(* IEC 61131-3 sources: daoli-st-library/DL_Base, 243 files *)

(* ---- E_DL_ControlModeSel.st ---- *)
// E_DL_ControlModeSel v1.0.0
// 开源溯源：AixOCAT / URL https://github.com/AixOCAT / 许可证 MIT / 借鉴 CONTROL_MODE 枚举语义（手/自动/停止三态），clean-room 重写
(*
  道莅工业代码库 | DL_Base | E_DL_ControlModeSel
  版本: 1.0.0 | 日期: 2026-11-23 | 轮次: R75
  功能: 手动/自动/停止三态控制模式枚举（strict 口径，配 MANUAL 覆写件族）
  邻件关系: 与 E_SMStatus 语义相邻（状态机状态 vs 操作模式选择），本件为
            模式选择属主；引用方（覆写/手自动切换族）只引用不重声明（R12）
  使用约定: 全库唯一属主，其他件引用时由 L2 闸按类型名自动回溯本文件；
            成员值固定步进 10，禁止中途插值改序（防历史引用漂移）
*)
TYPE E_DL_ControlModeSel :
(
    eManual := 0,    // 手动模式（操作员直控，联锁保留）/ Manual mode, operator direct with interlocks
    eAuto   := 10,   // 自动模式（程序/上位调度）/ Auto mode, program or supervisory driven
    eStop   := 20    // 停止模式（受控停机，输出回安全位）/ Stop mode, controlled stop to safe outputs
);
END_TYPE

(* ---- FB_DL_EStopMonitor.st ---- *)
(*==============================================================================
 * 组件名称 (Component)  : FB_DL_EStopMonitor
 * 所属子库 (Sublibrary) : DL_Base
 * 当前版本 (Version)    : 1.0.0
 * 兼容性   (Platform)   : CODESYS 3.5+ / TwinCAT 3 / 汇川 InoProShop / 施耐德 Machine Expert
 *                         仅依赖 Standard.library（TON / R_TRIG / F_TRIG / ABS），
 *                         零厂商私有库
 * 功能描述 (Function)   : 急停双通道监视：通道语义 TRUE=回路闭合（健康）。
 *                         任一通道断开 → bSafe 立即 FALSE（安全侧一级拦截，
 *                         不等确认窗）；两通道电平不一致（bCh1 <> bCh2）持续
 *                         tMismatchWin → bMismatch 锁存 + 首出通道号 eFirstOut
 *                         锁存（先断开的通道，F_TRIG 双实例竞争记录）；复位须
 *                         双通道恢复一致（bCh1 ∧ bCh2）且 bReset 上升沿才清
 *                         bMismatch/首出（规格指定）。
 * 接口     (Interface)  : 输入 bCh1 通道 1（TRUE=闭合健康）、bCh2 通道 2、
 *                         tMismatchWin 失配确认窗（域 > T#0S）、bReset 复位；
 *                         输出 bSafe 可运行判据（双通道健康 ∧ 无失配锁存）、
 *                         bMismatch 失配锁存、eFirstOut 首出通道号（锁存）、
 *                         eErrCode 错误码、bError 故障标志。
 * 边界     (Boundary)   : ① **属主边界（写死）：本件只做双通道监视判据，不切断
 *                         执行器、不做安全认证**（安全切断由安全继电器/IO 映射层
 *                         双保险执行，本件为诊断与允许运行判据源）。
 *                         ② 首出归因：双 F_TRIG 竞争窗口内先到沿者赢（同拍
 *                         双断时按 bCh1 优先判定，头注释声明：同拍双断无法区分
 *                         物理先后，eFirstOut 取 eCh1，规格允许的确定性归因）。
 *                         ③ 双通道同拍齐断（一致断开）不判失配：bSafe=FALSE
 *                         照常拦截，eFirstOut 保持 eNone（一致事件无失配语义）。
 *                         ④ 失配确认 TON 的 IN 派生式（bCh1 <> bCh2）∧ 通道
 *                         未齐断，段 0 无条件调用；出窗自复位（不一致消失即
 *                         复位，无外部沿清零依赖）。
 *                         ⑤ 锁存解除路径：bMismatch/eFirstOut 解除边 = 双通道
 *                         健康 ∧ bReset 上升沿（可达，头注释声明，R188/R152）。
 *                         ⑥ 零全局耦合（无 GVL / VAR_EXTERNAL / 物理地址）。
 * 分工声明 (Scope)      : 与 `FB_DL_RedundantSwitch` 分工：通道二选一归那件、
 *                         急停一致性监视归本件；与 `FB_DL_EdgeOrderCheck` 分工：
 *                         通用顺序校验归那件，本件首出归因为急停专用语义。
 * 来源标签 (Source Tag) : IEC 61131-3 标准语义的道莅防御性实现（双通道一致性
 *                         监视为标准安全监视语义）
 * 码表     (Codes)      : 本件不占用任何全局数字码位。出口为 BOOL 组 +
 *                         ENUM 通道号/错误码；数字码位待主控收口阶段统一派号。
 * 红线自检 (Redline)    : R1 ✓ 零 GVL/VAR_EXTERNAL ｜ R2 ✓ 零 %I/%Q/%M ｜ R3 ✓ 纯 IEC 61131-3
 *                         R4 ✓ 一级拦截不等窗 + 锁存解除可达 + 归因唯一 ｜ R5 ✓ 声明逐行同行双语注释
 *                         R6 ✓ ENUM 状态机不用（首出枚举 + 锁存态） ｜ R7 ✓ 一 TON 两 F_TRIG 一 R_TRIG 段 0 无条件刷新
 * 修订历史 (Revision)   : 2026-11-20  v1.0.0  R50 首版（批次 2 · 序号 10）
 * 验收向量 (Acceptance) : ① 双通道 TRUE，bCh1 在 t0 断开且 tMismatchWin 内未
 *                         恢复 → bMismatch=TRUE、eFirstOut=eCh1、bSafe=FALSE；
 *                         ② bCh1 断开 20ms 内恢复（tMismatchWin=100MS）→
 *                         tonMis 未到，bMismatch 保持 FALSE；③ 失配锁存后
 *                         bCh1/bCh2 均 TRUE + bReset 上升沿 → bMismatch=
 *                         FALSE、eFirstOut=eNone、bSafe=TRUE；④ 双通道同拍
 *                         齐断 → bSafe=FALSE，bMismatch=FALSE，eFirstOut=eNone。
 *==============================================================================*)

(*-----------------------------------------------------------------------------
 * 枚举: E_DL_EstChannel（首出通道号，锁存回放）
 *----------------------------------------------------------------------------*)
TYPE E_DL_EstChannel :
(
    eNone := 0,   // 无首出（未发生失配或同拍齐断） / No first-out
    eCh1  := 1,   // 首出通道 1 / First-out channel 1
    eCh2  := 2    // 首出通道 2 / First-out channel 2
);
END_TYPE

(*-----------------------------------------------------------------------------
 * 枚举: E_DL_EstErr（错误码；信息级不置 bError，故障级恒伴 bError=TRUE）
 *----------------------------------------------------------------------------*)
TYPE E_DL_EstErr :
(
    eOk      := 0,   // 正常 / Normal
    eCfgBad  := 1,   // 故障级：确认窗组态非法（<= T#0S） / Fault: window config illegal
    eMisLock := 2    // 故障级：失配锁存回放（归因见 eFirstOut） / Fault: mismatch latched replay
);
END_TYPE

FUNCTION_BLOCK FB_DL_EStopMonitor
VAR_INPUT
    bCh1         : BOOL := TRUE;    // 通道 1（TRUE=回路闭合健康） [-] / Channel 1, TRUE means healthy closed
    bCh2         : BOOL := TRUE;    // 通道 2（TRUE=回路闭合健康） [-] / Channel 2, TRUE means healthy closed
    tMismatchWin : TIME := T#100MS; // 失配确认窗，域 > T#0S [ms] / Mismatch confirmation window
    bReset       : BOOL := FALSE;   // 复位（须双通道健康后上升沿才生效） [-] / Reset, effective only with both channels healthy
END_VAR
VAR_OUTPUT
    bSafe     : BOOL;                // 可运行判据（双通道健康 ∧ 无失配锁存） [-] / Safe-to-run verdict
    bMismatch : BOOL;                // 失配锁存（解除 = 双通道健康 ∧ 复位沿） [-] / Mismatch latch
    eFirstOut : E_DL_EstChannel;     // 首出通道号（锁存回放，R189） / First-out channel, latched
    eErrCode  : E_DL_EstErr;         // 错误码出口 / Error code outlet
    bError    : BOOL;                // 故障标志（失配锁存或组态） [-] / Error flag
END_VAR
VAR
    _bMisLatch: BOOL;                // 失配锁存位（解除路径见头注释⑤） / Latched mismatch bit
    _eFirst   : E_DL_EstChannel := E_DL_EstChannel.eNone;   // 首出通道锁存 / Latched first-out channel
    _bCfgBad  : BOOL;                // 组态非法当拍量 [-] / Illegal configuration this scan
    _bCfgLatch: BOOL;                // 组态故障锁存位（解除沿 = 双通道健康 ∧ bReset 上升沿） / Latched config fault
    _bBothOk  : BOOL;                // 双通道健康当拍量 [-] / Both channels healthy
    rtReset   : R_TRIG;              // 复位沿实例，段 0 无条件调用 / Reset edge instance
    ftCh1     : F_TRIG;              // 通道 1 下降沿（断开）实例，段 0 无条件调用 / Ch1 falling-edge instance
    ftCh2     : F_TRIG;              // 通道 2 下降沿（断开）实例，段 0 无条件调用 / Ch2 falling-edge instance
    tonMis    : TON;                 // 失配确认窗，段 0 无条件调用 / Mismatch confirmation TON
END_VAR

(* —— 段 0：组态闸 + 全部沿/定时器无条件周期刷新（R6/R7） —— *)
_bCfgBad := (tMismatchWin <= T#0S);            // 确认窗域闸 / Window configuration gate
_bBothOk := bCh1 AND bCh2;                     // 双通道健康判据 / Both channels healthy
rtReset(CLK := bReset);                        // 复位沿，每拍必调 / Reset edge, every scan
ftCh1(CLK := bCh1);                            // 通道 1 断开沿，每拍必调 / Ch1 open edge, every scan
ftCh2(CLK := bCh2);                            // 通道 2 断开沿，每拍必调 / Ch2 open edge, every scan
tonMis(IN := (bCh1 <> bCh2) AND (NOT _bMisLatch) AND (NOT _bCfgLatch),
       PT := tMismatchWin);                    // 失配确认窗（出窗自复位：不一致消失即清，头注释④） / Mismatch window, self-resetting

(* —— 段 1：复位沿（须双通道健康才生效；清失配/首出/组态锁存） —— *)
IF rtReset.Q AND _bBothOk THEN
    _bMisLatch := FALSE;                       // 清失配锁存（可达解除路径，头注释⑤） / Clear mismatch latch
    _eFirst := E_DL_EstChannel.eNone;          // 清首出归因 / Clear first-out
    _bCfgLatch := FALSE;                       // 清组态锁存 / Clear config latch
END_IF
IF _bCfgBad AND (NOT _bCfgLatch) THEN
    _bCfgLatch := TRUE;                        // 组态锁存 / Latch config fault
END_IF

(* —— 段 2：首出归因（失配未锁存期，先断沿者赢；同拍双断 bCh1 优先，头注释②） —— *)
IF (NOT _bMisLatch) AND (bCh1 <> bCh2) THEN
    IF ftCh1.Q THEN
        _eFirst := E_DL_EstChannel.eCh1;       // 通道 1 先断归因 / Ch1 first-out
    ELSIF ftCh2.Q THEN
        _eFirst := E_DL_EstChannel.eCh2;       // 通道 2 先断归因 / Ch2 first-out
    END_IF
END_IF

(* —— 段 3：失配确认锁存（窗到锁存；同拍齐断不判失配，头注释③） —— *)
IF tonMis.Q AND (NOT _bMisLatch) THEN
    _bMisLatch := TRUE;                        // 失配锁存（R189：锁存回放，不在故障相重推断） / Latch mismatch
END_IF

(* —— 段 4：出口单点映射（名实双出口同源，R191） —— *)
bSafe := _bBothOk AND (NOT _bMisLatch) AND (NOT _bCfgLatch);   // 可运行判据（安全侧一级拦截不等窗） / Safe verdict, immediate intercept
bMismatch := _bMisLatch;                       // 失配出口 / Mismatch outlet
eFirstOut := _eFirst;                          // 首出出口 / First-out outlet
IF _bCfgLatch THEN
    bError := TRUE;                            // 故障标志（组态级，R45 配对） / Error flag
    eErrCode := E_DL_EstErr.eCfgBad;           // 组态故障码 / Config fault code
ELSIF _bMisLatch THEN
    bError := TRUE;                            // 故障标志（失配级） / Error flag
    eErrCode := E_DL_EstErr.eMisLock;          // 失配锁存回放码 / Mismatch replay code
ELSE
    bError := FALSE;                           // 正常 / Normal
    eErrCode := E_DL_EstErr.eOk;               // 正常码 / OK code
END_IF

END_FUNCTION_BLOCK

(* ---- FB_DL_FrequencyMeasure.st ---- *)
(*==============================================================================
 * 组件名称 (Component)  : FB_DL_FrequencyMeasure
 * 溯源说明 (Provenance): 道莅 clean-room 防御性实现（IEC 61131-3 纯净实现，闭源文档仅借语义，零代码行）
 * 所属子库 (Sublibrary) : DL_Base / Timing
 * 当前版本 (Version)    : 1.0.0
 * 兼容性   (Platform)   : CODESYS 3.5 / TwinCAT 3 / 汇川 InoProShop / 施耐德
 *                         Machine Expert；纯 IEC 61131-3（第 3 版），仅用
 *                         Standard.library 的 R_TRIG / TON / TIME_TO_REAL
 * 组件分类 (Category)   : 功能块（FUNCTION_BLOCK）· 门时计数测频
 * 功能一句话 (Summary)  : 用固定门时间数脉冲上升沿，算出外部脉冲的频率 [Hz]，
 *                         并把当拍分辨率与低频死区显式化。
 *
 * 本件存在的意义 (Why this unit exists)
 *   定时器族此前只有「生」没有「测」：PulseGenerator 生脉冲、SamplingTrigger
 *   生节拍、CycleTimeMeasure 测任务周期，**没有任何件测量外部脉冲频率**。
 *   脉冲流量计的 K 系数换算、编码器线速度、风机转速全部落在这一格。
 *   R21 已判「频率发生器不立」（与 PulseGenerator 重叠），但测量侧与之相反，
 *   是真实缺口：测频的不确定度、分辨率、低频死区必须显式给出，否则现场
 *   拿一个小数抖动值当转速用。
 *
 * 测量原理 (Principle)
 *   门时间内数上升沿：f = N / T_gate。分辨率 = 1 / T_gate（门越长分辨率越高、
 *   响应越慢，这是本件必须让调用方自己权衡的取舍，故做成引脚而非内部默认）。
 *   门到时立即发布、计数清零、重开门——不存在「测量间隙」的可配置语义，
 *   间隙固定为 1 个扫描周期（绝对时间不确定度见遗留假设）。
 *
 * 遗留假设 (Assumption) —— 测量不确定度，不得声称精确
 *   ① 门切换拍可能多计或漏计 **1 个沿**，故测量不确定度为 ±1 计数，
 *      折算 ±1/T_gate Hz。这是门时计数法的原理性下限，不是实现缺陷；
 *   ② 门时间以任务周期为量化单位，实际门时间 = 设定值 ± 1 个任务周期；
 *   ③ 分辨率引脚 fFreqRes 给出的是「当拍实际分辨率」= 1000 / 门毫秒数，
 *      调用方据此判断低频侧的可信度（低频 + 短门 → 分辨率极粗）；
 *   ④ 低于 fLowFreqDead 一律输出 0（信息 0465），不输出抖动小数冒充低频——
 *      停机的流量计输出 0.37 Hz 会让操作工以为还在流。
 *
 * 边界安全 (Boundary)
 *   ① tGateTime < T#1MS → 钳到 1 ms + 信息 0464；> T#10S → 钳到 10 s + 信息 0464；
 *   ② 门时间经钳位后为 0 属结构性不可达（防御纵深）→ 故障 03B4、回 eIdle；
 *   ③ 计数在门切换拍出现回退（外部改写或溢出）→ 故障 03B5、bValid = FALSE，
 *      并丢弃本门计数从零重开门（本件无复位引脚，故为自愈式处理，见实现注释）；
 *   ④ R_TRIG 与 TON 实例在主体最前部**无条件刷新**（R40 家族），门重启经
 *      「断输入一拍」标志 _bGateBreak 实现，调用后立即自清；
 *   ⑤ CASE 落 ELSE 置 03B5 并回 eIdle（非法状态兜底，与③共用一码，R90）。
 * 节律 (Cycle order)
 *   段 1 每拍预置 → 段 2 首扫初始化 → 段 3 参数钳位 → 段 4 边沿与定时器无条件
 *   刷新（含计数累加）→ 段 5 计数回退检测 → 段 6 状态机（只做迁移）→
 *   段 7 发布（eReady 相内单拍，唯一写入点）→ 段 8 迁移收尾 → 段 9 出口。
 *
 * 错误码    : 16#0001_0464 门时间越界已钳位到 1 ms~10 s——信息级，正常防御
 *             16#0001_0465 频率低于死区，已按 0 输出——信息级，不输出抖动小数
 *             16#0001_03B4 门时间钳位后仍非法（为 0），无法测频——故障级，bValid = FALSE
 *             16#0001_03B5 门内计数回退不可信（含状态机 ELSE 兜底复用，R90）——故障级
 *             16#0001_03B6 预留禁用（故障级，不得挪用）
 * 码位总账  : 16#0001_0464 用 / 16#0001_0465 用 ｜ 16#0001_03B4 用 / 16#0001_03B5 用 / 16#0001_03B6 预留
 * 状态机    : E_DL_FreqMeasState（eIdle / eGating / eReady / eFault），CASE 含 ELSE
 *             兜底，ELSE 分支置 16#0001_03B5 并回 eIdle；失能无条件回 eIdle
 * 采样约定  : 每任务周期调用一次；门时间由 tGateTime 给定，不读系统时钟
 * 依赖说明  : 无 DL_ 内部依赖；仅 Standard.library 的 R_TRIG / TON / TIME_TO_REAL
 * 验收向量  : V1 100 ms 门、1 kHz 脉冲 → fFreq ≈ 100.0，fFreqRes = 10.0，bValid = TRUE
 *             V2 100 ms 门、0.2 Hz 脉冲（死区内）→ fFreq = 0，eErr = 0465，bValid = TRUE
 *             V3 门时间 0 ms → 钳到 1 ms 且 eErr = 0464，仍返回测量（钳位主向量）
 *             V4 门时间 20 s → 钳到 10 s 且 eErr = 0464
 *             V5 门切换拍清零后立刻被外部写回大值（构造计数回退）→ eErr = 03B5，
 *                bValid = FALSE，随后自愈重开（R40 跨相主向量）
 *             V6 失能 → eIdle，bValid = FALSE，fFreq 保持末次值不跳变（恢复首拍不阶跃）
 * 红线自检  : 全局变量声明零使用 / 外部变量访问零使用 / 物理地址零使用 ｜ 纯 IEC 61131-3 ｜ 除法前置
 *             判零（门时恒 ≥ 1 ms，构造性非零，另设显式闸门）｜ 浮点比较只用
 *             容差与大小比较，无判等 ｜ 循环无、计数带上界饱和 ｜ 全变量双语
 *             同行注释 ｜ ENUM + CASE 含 ELSE ｜ R_TRIG / TON 在主体最前部无条件
 *             刷新 ｜ 无魔法数
 * 修订历史  : 2026-11-16  v1.0.0  首版入库（R22 · 批 1 · 定时器族第五轴）
 *============================================================================*)

(*-----------------------------------------------------------------------------
 * 枚举: E_DL_FreqMeasState（归属本功能块，同文件发布，全库唯一定义）
 * 含义: 门时测频的离散相位。0 起步长 10，便于后续插态。
 *-----------------------------------------------------------------------------*)
TYPE E_DL_FreqMeasState :
(
    eIdle     := 0,    // 待机：未使能或门时间非法 / Idle, disabled or gate time illegal
    eGating   := 10,   // 计数中：门时间内数上升沿 / Gating, counting rising edges inside the gate
    eReady    := 20,   // 发布相：门到后单拍发布并重开 / Ready, one scan to publish then reopen
    eFault    := 99    // 故障：门时间非法，待参数恢复 / Fault, gate time illegal until it recovers
);
END_TYPE

FUNCTION_BLOCK FB_DL_FrequencyMeasure
VAR_INPUT
    bPulse       : BOOL;                       // 待测脉冲，任意占空比 / pulse under test, any duty cycle
    bEnable      : BOOL;                       // 使能，FALSE 时停止计数并回待机 / enable, FALSE stops counting and returns to idle
    tGateTime    : TIME := T#100MS;            // 门时间 [ms]，范围 1~10000 / gate time [ms], range 1~10000
    fLowFreqDead : REAL := 0.5;                // 低频死区 [Hz]，低于此值输出 0 / low frequency dead band [Hz], output zero below it
END_VAR
VAR_OUTPUT
    fFreq        : REAL;                       // 测量频率 [Hz]，分辨率 1/tGateTime / measured frequency [Hz], resolution 1/gate time
    fFreqRes     : REAL;                       // 当拍实际分辨率 [Hz] / actual resolution of the current scan [Hz]
    uLastCount   : UDINT;                      // 上一门内上升沿个数 [个] / rising edge count of the previous gate
    bValid       : BOOL;                       // 输出可用标志 / outputs usable flag
    eErr         : UDINT;                      // 错误码，0 表示无错 / error code, 0 means no error
    bError       : BOOL;                       // 故障级标志，仅故障级错误置位 / fault-class flag, set only on fault-level codes
END_VAR
VAR
    fbEdge       : R_TRIG;                     // 脉冲上升沿检测，段 4 无条件刷新 / pulse rising edge detector, refreshed unconditionally
    fbGate       : TON;                        // 门时间计时，段 4 无条件刷新 [ms] / gate timer, refreshed unconditionally
    _eState      : E_DL_FreqMeasState := E_DL_FreqMeasState.eIdle; // 当前相位 / current phase
    _bInit       : BOOL := FALSE;              // 首扫标志，初值 FALSE 取非判定 / first-scan flag, FALSE initialised and tested negated
    _tGateUse    : TIME := T#100MS;            // 生效门时间 [ms]，已钳位 / effective gate time after clamping
    _fDeadUse    : REAL := 0.5;                // 生效低频死区 [Hz]，已钳位 / effective dead band after clamping
    _uCount      : UDINT;                      // 本门内上升沿累计 [个] / rising edges accumulated inside the current gate
    _uCountPrev  : UDINT;                      // 上拍计数快照，唯一写入点在段 9 [个] / previous-scan count snapshot, single write point
    _uLastCountH : UDINT;                      // 上一门计数保持量 [个] / held edge count of the previous gate
    _fFreqHeld   : REAL;                       // 频率保持量 [Hz] / held frequency
    _fResHeld    : REAL;                       // 分辨率保持量 [Hz] / held resolution
    _bHaveMeas   : BOOL;                       // 是否已完成过一次测量 / whether one full measurement has completed
    _bGateBreak  : BOOL;                       // 门计时器断输入一拍标志 / gate timer one-scan break flag
    _bParamFault : BOOL;                       // 门时间参数非法标志 / gate time illegal flag
    _bRollback   : BOOL;                       // 计数回退标志 / counter rollback flag
    _fGateMs     : REAL;                       // 门时间毫秒数 [ms]，用于换算 / gate time in milliseconds used by the conversions
END_VAR
VAR CONSTANT
    DL_GATE_MIN_MS  : DINT := 1;               // 门时间下限 [ms] / gate time floor [ms]
    DL_GATE_MAX_MS  : DINT := 10000;           // 门时间上限 [ms] / gate time ceiling [ms]
    DL_TIME_ZERO    : TIME := T#0MS;           // 时间零值基准 [ms] / time zero reference
    DL_MS_PER_S     : REAL := 1000.0;          // 毫秒与秒的换算系数 [ms/s] / milliseconds per second
    DL_CNT_MAX      : UDINT := 16#FFFF_FFFF;   // 计数饱和上界 [个]，不回绕 / counter saturation ceiling, never wraps
    DL_DEAD_MAX     : REAL := 1000.0;          // 死区参数上限 [Hz]，防超界 / dead band parameter ceiling [Hz]
    DL_DEAD_MIN     : REAL := 0.0;             // 死区参数下限 [Hz]，负值无意义 / dead band parameter floor [Hz]
END_VAR

(*------------------------------------------------------------------------------
 * 段 1｜每拍预置（状态量与保持量不预置，输出在段 9 单点写入）
 *      Per-scan presets, held values and outputs are untouched here
 *-----------------------------------------------------------------------------*)
eErr         := 16#0000_0000;                  // 错误码每拍重算 / error code recomputed every scan
bError       := FALSE;                         // 故障标志每拍重算 / fault flag recomputed every scan
bValid       := FALSE;                         // 可用标志每拍重算 / usable flag recomputed every scan
_bParamFault := FALSE;                         // 参数非法标志预清零 / parameter fault flag pre-cleared
_bRollback   := FALSE;                         // 回退标志预清零 / rollback flag pre-cleared

(*------------------------------------------------------------------------------
 * 段 2｜首扫初始化（R19：bInit 初值 FALSE，判据取非）
 *      First-scan initialisation
 *-----------------------------------------------------------------------------*)
IF NOT _bInit THEN
    _eState     := E_DL_FreqMeasState.eIdle;   // 相位待机 / phase idle
    _uCount     := 0;                          // 计数清零 / counter cleared
    _uCountPrev := 0;                          // 快照清零 / snapshot cleared
    _uLastCountH := 0;                         // 上一门计数清零 / previous gate count cleared
    _fFreqHeld  := 0.0;                        // 频率保持量清零 / held frequency cleared
    _fResHeld   := 0.0;                        // 分辨率保持量清零 / held resolution cleared
    _bHaveMeas  := FALSE;                      // 尚无测量 / no measurement yet
    _bGateBreak := TRUE;                       // 首个门从零开始计时 / the first gate starts from zero
    _bInit      := TRUE;                       // 首扫只做一次 / the first scan runs once
END_IF

(*------------------------------------------------------------------------------
 * 段 3｜参数钳位（门时间 1 ms~10 s；死区 0~上限）
 *      Parameter clamping, gate time one millisecond to ten seconds
 *-----------------------------------------------------------------------------*)
IF TIME_TO_DINT(tGateTime) < DL_GATE_MIN_MS THEN
    _tGateUse := DINT_TO_TIME(DL_GATE_MIN_MS); // 钳到下限 1 ms / clamped to the floor
    eErr      := 16#0001_0464;                 // 信息级：门时间已钳位 / informational: gate time clamped
ELSIF TIME_TO_DINT(tGateTime) > DL_GATE_MAX_MS THEN
    _tGateUse := DINT_TO_TIME(DL_GATE_MAX_MS); // 钳到上限 10 s / clamped to the ceiling
    eErr      := 16#0001_0464;                 // 信息级：门时间已钳位 / informational: gate time clamped
ELSE
    _tGateUse := tGateTime;                    // 域内直通 / passed through inside the domain
END_IF

(* 钳位后仍为 0：结构性不可达，保留 03B4 给「门时间为 0 的构造路径」（防御纵深） *)
(* Still zero after clamping is structurally unreachable, kept as defense in depth *)
IF _tGateUse <= DL_TIME_ZERO THEN
    _tGateUse    := DINT_TO_TIME(DL_GATE_MIN_MS); // 兜底回 1 ms，防后续除零 / fallback to one millisecond, no division by zero downstream
    _bParamFault := TRUE;                      // 参数故障标志 / parameter fault flag
    eErr         := 16#0001_03B4;              // 故障级：门时间非法 / fault: illegal gate time
    bError       := TRUE;                      // 置故障标志 / raise the fault flag
END_IF

_fDeadUse := LIMIT(DL_DEAD_MIN, fLowFreqDead, DL_DEAD_MAX); // 死区钳进 0~1000 Hz / dead band clamped

(*------------------------------------------------------------------------------
 * 段 4｜边沿与定时器无条件刷新（R40：一律在 CASE 之外、每拍必调）
 *      Edge detector and timer refreshed unconditionally, outside the CASE
 *-----------------------------------------------------------------------------*)
fbEdge(CLK := bPulse);                          // 脉冲沿无条件刷新 / pulse edge refreshed unconditionally

IF fbEdge.Q AND (_eState = E_DL_FreqMeasState.eGating) THEN
    IF _uCount < DL_CNT_MAX THEN
        _uCount := _uCount + 1;                 // 门内计数，饱和不回绕 / counted inside the gate, saturating
    END_IF
END_IF

fbGate(IN := bEnable AND (_eState = E_DL_FreqMeasState.eGating) AND (NOT _bGateBreak),
       PT := _tGateUse);                        // 门计时无条件刷新 / gate timer refreshed unconditionally
_bGateBreak := FALSE;                           // 断输入拍在调用后自清（R40 自清位置） / break self-cleared right after the call

(*------------------------------------------------------------------------------
 * 段 5｜计数回退检测（本件无复位引脚，故为自愈式：弃本门、从零重开）
 *      Counter rollback detection, self-healing because there is no reset pin
 *-----------------------------------------------------------------------------*)
IF _uCount < _uCountPrev THEN
    _bRollback := TRUE;                         // 标记回退 / rollback flagged
    _uCount    := 0;                            // 丢弃不可信计数 / drop the untrustworthy count
    _bGateBreak := TRUE;                        // 门计时从零重启 / gate timer restarted from zero
    _eState    := E_DL_FreqMeasState.eIdle;     // 回待机，下一拍重新开门 / back to idle, the gate reopens next scan
    eErr       := 16#0001_03B5;                 // 故障级：计数回退不可信 / fault: counter rollback, untrustworthy
    bError     := TRUE;                         // 置故障标志 / raise the fault flag
END_IF

(*------------------------------------------------------------------------------
 * 段 6｜相位机（只做迁移，不写保持量；ELSE 兜底置 03B5 并回 eIdle）
 *      Phase machine, transitions only, a trailing ELSE falls back to 03B5 and idle
 *-----------------------------------------------------------------------------*)
CASE _eState OF

    E_DL_FreqMeasState.eIdle:                   // 待机：参数合法且使能即开门
        IF _bParamFault THEN
            _eState := E_DL_FreqMeasState.eFault; // 参数非法转故障 / illegal parameters go to fault
        ELSIF bEnable THEN
            _uCount    := 0;                    // 新门从零计数 / a new gate starts at zero
            _bGateBreak := TRUE;                // 门计时从零开始 / gate timer starts from zero
            _eState    := E_DL_FreqMeasState.eGating; // 进计数相 / enter the gating phase
        END_IF

    E_DL_FreqMeasState.eGating:                 // 计数中：门到即转发布相
        IF NOT bEnable THEN
            _eState := E_DL_FreqMeasState.eIdle; // 失能回待机 / disabled, back to idle
        ELSIF fbGate.Q THEN
            _eState := E_DL_FreqMeasState.eReady; // 门到，转发布相（发布在段 7） / gate done, publishing happens in segment seven
        END_IF

    E_DL_FreqMeasState.eReady:                  // 发布相：段 7 发布、段 8 迁移
        IF NOT bEnable THEN
            _eState := E_DL_FreqMeasState.eIdle; // 失能中止 / disabled, abort
        END_IF

    E_DL_FreqMeasState.eFault:                  // 故障：参数恢复即回待机
        IF NOT _bParamFault THEN
            _eState := E_DL_FreqMeasState.eIdle; // 参数已恢复 / parameters recovered
        END_IF

    ELSE
        eErr    := 16#0001_03B5;                // 兜底复用：非法状态（R90 不加码） / fallback reuse: illegal state
        bError  := TRUE;                        // 置故障标志 / raise the fault flag
        _uCount := 0;                           // 计数清零，绝不带着脏计数继续 / counter cleared, never continue with a dirty count
        _bGateBreak := TRUE;                    // 门计时重启 / gate timer restarted
        _eState := E_DL_FreqMeasState.eIdle;    // 回安全态 / back to the safe state
END_CASE

(*------------------------------------------------------------------------------
 * 段 7｜发布（eReady 相内单拍；fFreq / fFreqRes / uLastCount 的唯一写入点）
 *      Publish inside the ready phase, the single write point for all three values
 *-----------------------------------------------------------------------------*)
IF _eState = E_DL_FreqMeasState.eReady THEN
    _fGateMs := TIME_TO_REAL(_tGateUse);        // 门时间换算为毫秒数 [ms] / gate time in milliseconds

    IF _fGateMs <= 0.0 THEN
        _fGateMs := DL_MS_PER_S;                // 除零兜底：结构性不可达 / division fallback, structurally unreachable
    END_IF

    _uLastCountH := _uCount;                    // 锁存本门计数 [个] / latch this gate count
    _fFreqHeld   := (UDINT_TO_REAL(_uLastCountH) / _fGateMs) * DL_MS_PER_S; // N/ms×1000 = N/s [Hz] / edges per millisecond to hertz
    _fResHeld    := DL_MS_PER_S / _fGateMs;     // 分辨率 = 1/T_gate [Hz] / resolution is one over the gate time

    IF _fFreqHeld < _fDeadUse THEN
        _fFreqHeld := 0.0;                      // 死区内输出 0，不输出抖动小数 [Hz] / inside the dead band output zero
        eErr       := 16#0001_0465;             // 信息级：低于死区按 0 输出 / informational: below the dead band, zero output
    END_IF

    _bHaveMeas := TRUE;                         // 已有一次完整测量 / one full measurement exists
    _uCount    := 0;                            // 计数清零，准备下一门 / counter cleared for the next gate
    _bGateBreak := TRUE;                        // 门计时从零重启 / gate timer restarted from zero
END_IF

(*------------------------------------------------------------------------------
 * 段 8｜迁移收尾（发布之后才允许 eReady → eGating，顺序不可反）
 *      Advance from ready back to gating only after the publish
 *-----------------------------------------------------------------------------*)
IF _eState = E_DL_FreqMeasState.eReady THEN
    _eState := E_DL_FreqMeasState.eGating;      // 回计数相 / back to the gating phase
END_IF

(*------------------------------------------------------------------------------
 * 段 9｜出口单点写入与可用性仲裁
 *      Single write point of the outputs and the usability arbitration
 *-----------------------------------------------------------------------------*)
fFreq      := _fFreqHeld;                       // 频率出口 [Hz] / frequency outlet
fFreqRes   := _fResHeld;                        // 分辨率出口 [Hz] / resolution outlet
uLastCount := _uLastCountH;                     // 上一门计数出口 [个] / previous gate count outlet
_uCountPrev := _uCount;                         // 快照在段末唯一写入（R45②） / snapshot written once at the end

IF bError THEN
    bValid := FALSE;                            // 故障级：输出不可用 / fault: outputs unusable
ELSIF NOT bEnable THEN
    bValid := FALSE;                            // 失能：输出不可用（值仍保持，供停机前趋势） / disabled: unusable, values still held
ELSE
    bValid := _bHaveMeas;                       // 已有完整测量才宣称可用 / usable only after a full measurement
END_IF

END_FUNCTION_BLOCK

(* ---- FB_DL_InterlockBypassAudit.st ---- *)
(*==============================================================================
 * 组件名称 (Component)  : FB_DL_InterlockBypassAudit
 * 所属子库 (Sublibrary) : DL_Base
 * 当前版本 (Version)    : 1.0.1
 * 兼容性   (Platform)   : CODESYS 3.5 / TwinCAT 3 / 汇川 InoProShop / Machine Expert
 *                         仅依赖 Standard.library（TON / R_TRIG），零厂商方言
 * 来源标签 (Source)     : t2-8-isa182（ISA-182 旁路管理方法论，clean-room 编写）
 * 功能描述 (Function)   : 联锁旁路全生命周期审计：申请沿进入旁路态并启动时限窗，
 *                         时限到期自动恢复并置信息级码；人工解除沿即时恢复。
 *                         申请沿 / 解除沿 / 超时到期三类事件写入 8 条深度环形台账，
 *                         台账带全局序号与旁路计数（饱和不回绕）。
 *                         旁路期间目标联锁位仍照常计算，仅放行判定被旁路——
 *                         放行判定归调用方按 bBypassActive 组合，本件不替代联锁本体。
 * 分工互引 (Boundary)   : 联锁本体的条件求值与首因锁存归 FB_DL_InterlockMatrix；
 *                         安全门的旁路申请登记归 FB_DL_SafetyDoorAuditBank；
 *                         本件只负责旁路时限与事件台账审计，三者互不替代。
 * 边界与语义披露 (Boundary disclosure) :
 *   1) 时限窗 tBypassWindow <= T#0S 视为组态非法：置故障级码并拒绝进入旁路态，
 *      已在旁路态的不受影响（组态变更不追溯已生效旁路），故障锁存经复位沿清除。
 *   2) 同拍「申请沿 + 解除沿」：解除优先（安全侧）——旁路不进入、不记申请事件。
 *   3) 旁路态不锁存联锁故障：本件是审计器不是联锁本体，故障锁存语义归联锁件。
 *   4) 台账为 8 条环形，写满后覆盖最旧条目并置信息级提示；写指针回卷由模运算
 *      等价的显式 IF 归零实现，不做越界写。
 *   5) 旁路计数为 USINT 饱和计数：255 + 1 停在 255 不回绕；计数顶格本身可由
 *      uBypassCount = 255 直接观测，故不另设码位（R90 反证成立，不加码）。
 * 故障码表 (Error codes) :
 *   16#0001_03EE [故障级] 时限窗组态非法（<= T#0S），拒绝进入旁路态
 *                 反证：该场景仅可由「申请沿被拒 + 状态停 eIdle」观测，但拒因
 *                 （时限非法还是使能关闭）不可区分，现有输出组合无法唯一还原。
 *   16#0001_04B1 [信息级] 时限到期自动恢复（旁路被时限收割）
 *                 反证：到期恢复与人工解除对外都表现为退出旁路态，唯一差异
 *                 是台账事件种类，无码时 HMI 无法区分两类恢复事件。
 *                 回落路径（v1.0.1 · L1）：下一轮旁路申请被受理时归零——
 *                 该事件码只描述「上一轮的收割事实」，新一轮开始即不再是当下事件。
 *   16#0001_04B2 [信息级] 台账环形已回卷（最旧条目被覆盖，审计完整性降级）
 *                 反证：回卷后 nLedgerCount 恒为 8，与「恰好写满未回卷」的
 *                 输出组合完全相同，不可由现有输出观测。
 *                 回落路径（v1.0.1 · L1）：一次性事件码（bWrapCoded 单次置位），
 *                 复位沿清除；回卷状态本身由 bLedgerWrapped 常驻表达（状态与
 *                 事件分离：码承载事件，位承载状态）。
 *   非法状态拦截复用全库惯用码 16#0001_0005（不新占号）。
 * 码位总账 (Code ledger) : 16#0001_03EE 用 ｜ 16#0001_04B1 用 / 16#0001_04B2 用
 * 依赖     (Depends)    : 无 DL_ 内部依赖；Standard.library: TON / R_TRIG
 * 红线自检 (Redline)    : R1 ✓ 零全局变量与 VAR_EXTERNAL ｜ R2 ✓ 零 %I/%Q 物理地址
 *                         R3 ✓ 纯 IEC 61131-3 标准库 ｜ R4 ✓ 时间窗判零 / 计数饱和 / 指针无涉
 *                         R5 ✓ 全变量中英双语同行注释 ｜ R6 ✓ 三态 ENUM + CASE + ELSE 兜底
 *                         R7 ✓ 一沿三实例主体最前部无条件刷新
 * 修订历史 (Revision)   :
 *   2026-11-22  v1.0.0  首版入库（R68 构建轮 · 批 1 · 目标 1）
 *   2026-11-22  v1.0.1  R69 点修①：迁相（组态故障打断 / 非法态兜底）补 bBypassOn := FALSE，
 *                       防新组态首旁路立即到期；点修⑤：信息码 04B1 随新一轮旁路受理回落、
 *                       04B2 改一次性事件码并由复位沿回落（回卷状态仍由 bLedgerWrapped 常驻）
 *============================================================================*)

(*-----------------------------------------------------------------------------
 * 枚举: E_DL_BypassState（归属 DL_Base，与 FB_DL_InterlockBypassAudit 同文件）
 * 含义: 旁路审计主状态。数值步长留空位便于后续插态而不破坏已有工程。
 *----------------------------------------------------------------------------*)
TYPE E_DL_BypassState :
(
    eIdle     := 0,    // 未旁路：联锁照常生效 / No bypass, interlock fully effective
    eBypassed := 10,   // 旁路生效中：时限窗计时 / Bypass active, time window running
    eFault    := 99    // 组态故障：时限窗非法，拒绝一切新旁路 / Config fault, window illegal
);
END_TYPE

(*-----------------------------------------------------------------------------
 * 枚举: E_DL_BypassEventKind（归属 DL_Base，与 FB_DL_InterlockBypassAudit 同文件）
 * 含义: 台账事件种类，三类全生命周期事件一一对应。
 *----------------------------------------------------------------------------*)
TYPE E_DL_BypassEventKind :
(
    eNone   := 0,    // 无事件（台账空槽哨兵）/ No event, empty ledger slot sentinel
    eApply  := 1,    // 申请沿：进入旁路态 / Apply edge: bypass entered
    eReleaseByCmd     := 2,  // 解除沿：人工解除 / Release edge: manual release
    eReleaseByTimeout := 3   // 超时到期：自动恢复 / Timeout expiry: auto restore
);
END_TYPE

(*==============================================================================
 * 功能块: FB_DL_InterlockBypassAudit
 * 调用约定: 每个扫描周期无条件调用一次；申请沿与解除沿均为单拍沿语义。
 * 无状态泄漏: 全部状态驻留于实例私有 VAR，零全局引用，可多机组并行实例化。
 *============================================================================*)
FUNCTION_BLOCK FB_DL_InterlockBypassAudit
VAR_INPUT
    bBypassReq     : BOOL;                    // 旁路申请，上升沿生效 / Bypass request, rising edge
    bBypassRelease : BOOL;                    // 旁路解除，上升沿生效 / Bypass release, rising edge
    uInterlockId   : UINT  := 0;              // 目标联锁号 [号]，随事件入台账 / Target interlock id, logged per event
    uSourceId      : UINT  := 0;              // 申请源标识 [号]，随事件入台账 / Request source id, logged per event
    tBypassWindow  : TIME  := T#30S;          // 旁路时限窗 [s]，<= T#0S 组态非法 / Bypass window [s], <= 0 illegal
    bEnable        : BOOL  := TRUE;           // 审计使能，FALSE 时冻结不受理新申请 / Audit enable, FALSE freezes new requests
    bReset         : BOOL;                    // 上升沿：清除组态故障锁存 / Rising edge: clear config fault latch
END_VAR
VAR_OUTPUT
    bBypassActive  : BOOL;                   // 旁路生效中（供调用方放行判定组合）/ Bypass active for the caller gating
    uBypassCount   : USINT;                  // 累计旁路次数 [次]，255 饱和 / Total bypass count, saturates at 255
    nLedgerCount   : INT;                    // 台账有效条数 [条]，0..8 / Valid ledger entries, 0..8
    bLedgerWrapped : BOOL;                   // 台账已回卷覆盖（信息级）/ Ledger wrapped, oldest overwritten
    eLastEvent     : E_DL_BypassEventKind;   // 最近一次事件种类 / Kind of the most recent event
    uLastEventSeq  : UDINT;                  // 最近事件全局序号 [号] / Global sequence of the last event
    uLastTarget    : UINT;                   // 最近事件目标联锁号 [号] / Target id of the last event
    uLastSource    : UINT;                   // 最近事件申请源标识 [号] / Source id of the last event
    aLedgerKind    : ARRAY[0..7] OF E_DL_BypassEventKind; // 台账事件种类环形副本 / Ledger kind ring copy
    auLedgerTarget : ARRAY[0..7] OF UINT;    // 台账目标联锁号环形副本 / Ledger target ring copy
    auLedgerSource : ARRAY[0..7] OF UINT;    // 台账申请源标识环形副本 / Ledger source ring copy
    bError         : BOOL;                   // 故障标志（组态类锁存）/ Fault flag, configuration class latched
    uErrorId       : UDINT;                  // 故障码，0 = 无故障 / Error code, 0 = none
    eState         : E_DL_BypassState;       // 当前状态（供 HMI 诊断）/ Current state for HMI diagnosis
END_VAR
VAR
    fbTrigReq      : R_TRIG;                 // 申请沿检测实例 / Request edge detector
    fbTrigRel      : R_TRIG;                 // 解除沿检测实例 / Release edge detector
    fbTrigReset    : R_TRIG;                 // 复位沿检测实例 / Reset edge detector
    tonWindow      : TON;                    // 旁路时限窗计时实例 / Bypass window timer
    eStateInt      : E_DL_BypassState;       // 主状态机内部当前态 / Internal state machine state
    bWindowInvalid : BOOL;                   // 本拍时限窗组态非法 / Window config illegal this scan
    bConfigLatch   : BOOL;                   // 组态故障锁存（复位沿清除）/ Config fault latch, cleared by reset edge
    bBypassOn      : BOOL;                   // 旁路窗计时进行中（TON 的 IN 派生量）/ Window timing active, drives TON.IN
    aeKindInt      : ARRAY[0..7] OF E_DL_BypassEventKind; // 台账事件种类（内部）/ Ledger kind ring, internal
    auiTargetInt   : ARRAY[0..7] OF UINT;    // 台账目标联锁号（内部）/ Ledger target ring, internal
    auiSourceInt   : ARRAY[0..7] OF UINT;    // 台账申请源标识（内部）/ Ledger source ring, internal
    nWriteIdx      : INT;                    // 台账写指针 [0..7] / Ledger write pointer
    uEventTotal    : UDINT;                  // 累计事件总数 [件]，环形深度之外的真值 / Total events ever, truth beyond ring depth
    uSeqCounter    : UDINT;                  // 全局序号计数器 [号]，饱和 / Global sequence counter, saturating
    uCntInt        : USINT;                  // 旁路计数内部副本（饱和）/ Internal bypass counter, saturating
    uTargetInt     : UINT;                   // 最近事件目标号内部副本 / Internal copy of last target id
    uSourceInt     : UINT;                   // 最近事件源号内部副本 / Internal copy of last source id
    eLastEventInt  : E_DL_BypassEventKind;   // 最近事件种类内部副本 / Internal copy of last event kind
    uLastSeqInt    : UDINT;                  // 最近事件序号内部副本 / Internal copy of last event sequence
    bErrorInt      : BOOL;                   // 本拍故障置位累加（出口归并）/ Fault set accumulator of this scan
    bWrapCoded     : BOOL;                   // 回卷事件码已发标志（防每拍重发，复位沿撤销）/ Wrap event already coded, cleared by reset
    bFirstScan     : BOOL := TRUE;           // 上电首扫标志 / First-scan flag
END_VAR
VAR CONSTANT
    DL_BYP_RING_DEPTH : INT   := 8;            // 台账环形深度 [条]，与数组维度一致 / Ledger ring depth, matches arrays
    DL_BYP_CNT_MAX    : USINT := 255;          // 旁路计数饱和值 [次] / Bypass counter saturation
    DL_BYP_SEQ_MAX    : UDINT := 16#FFFF_FFFE; // 序号计数饱和值 [号] / Sequence counter saturation
    DL_BYP_IDX_NONE   : INT   := 0;            // 空槽哨兵：0 号槽事件种类 eNone / Empty slot via kind sentinel
END_VAR

(*------------------------------------------------------------------------------
 * 段 1｜无条件刷新区（红线 R7）：三沿 + 一计时，全部位于主体最前部
 *      Unconditional refresh zone: three edges and one timer at the very top
 *      TON 的 IN 用内部派生量 bBypassOn（旁路态驻留标志），禁挂外部引脚原值
 *-----------------------------------------------------------------------------*)
fbTrigReq(CLK := bBypassReq);
fbTrigRel(CLK := bBypassRelease);
fbTrigReset(CLK := bReset);
tonWindow(IN := bBypassOn, PT := tBypassWindow);

(*------------------------------------------------------------------------------
 * 段 2｜上电首扫（FB50-2①）：台账槽位显式落哨兵，不依赖默认零的巧合
 *      First-scan init: ledger slots forced to sentinels explicitly
 *-----------------------------------------------------------------------------*)
IF bFirstScan THEN
    FOR nWriteIdx := 0 TO (DL_BYP_RING_DEPTH - 1) DO
        aeKindInt[nWriteIdx] := E_DL_BypassEventKind.eNone;   // 空槽哨兵 / Empty slot sentinel
    END_FOR
    nWriteIdx   := 0;
    uEventTotal := 0;
    uSeqCounter := 0;
    uCntInt     := 0;
    bWrapCoded  := FALSE;   // 回卷事件码首扫未发 / Wrap event not yet coded
    eStateInt   := E_DL_BypassState.eIdle;
    bFirstScan  := FALSE;
END_IF

(*------------------------------------------------------------------------------
 * 段 3｜每拍预清（FB32-1：只准含单拍标志，禁入快照 / 累计 / 锁存量）
 *      Per-scan preset: single-scan flags only, no snapshots or latches
 *-----------------------------------------------------------------------------*)
bErrorInt := FALSE;

(*------------------------------------------------------------------------------
 * 段 4｜组态域闸（R151）：时限窗 <= T#0S 即非法；非法即锁存，复位沿 + 组态恢复可解除
 *      Config gate: window <= 0 is illegal; latched, cleared by reset edge with valid config
 *      解除路径自证：bReset 上升沿 AND 组态已改对（R152 可达性）
 *-----------------------------------------------------------------------------*)
bWindowInvalid := (tBypassWindow <= T#0S);

IF bWindowInvalid THEN
    bConfigLatch := TRUE;
END_IF

IF bConfigLatch THEN
    uErrorId  := 16#0001_03EE;   // 故障级：时限窗组态非法 / Fault: window config illegal
    bErrorInt := TRUE;           // R45 配对：故障码 3 行内置位 / Paired with the fault code
    eStateInt := E_DL_BypassState.eFault;
    (* R69 点修①（迁相补清）：故障打断旁路时同步撤窗计时量。原实现只迁相不清
     * bBypassOn，TON.IN 常真 -> 时限窗在故障期照走并在修复后率先到期，
     * 新组态首旁路一进 eBypassed 即被 tonWindow.Q 收割（04B1 误报、旁路退化）。 *)
    (* Phase migration also drops the window timing quantity, so the window cannot expire during the fault *)
    bBypassOn := FALSE;          // 迁相即断计时：TON.IN 归假 / Timing quantity dropped on migration
END_IF

(*------------------------------------------------------------------------------
 * 段 5｜主状态机（红线 R6）：ENUM + CASE + ELSE 兜底
 *      Main state machine with the mandatory ELSE fallback
 *      使能冻结语义：空闲相受理判据内串 bEnable，失能即拒绝新申请（不另设覆盖段，
 *      避免「禁用覆盖吃掉沿」类 R39 失真）；已生效旁路的时限窗照走（审计不中断）。
 *      同拍竞态（R275）：eBypassed 相内先消化解除沿，再消化超时迁移
 *-----------------------------------------------------------------------------*)
CASE eStateInt OF

    E_DL_BypassState.eIdle:
        (* 同拍「申请 + 解除」：解除优先（安全侧），申请沿作废不记台账 *)
        (* Same-scan request plus release: release wins on the safe side *)
        IF bEnable AND (NOT bConfigLatch) AND fbTrigReq.Q AND (NOT fbTrigRel.Q) THEN
            uErrorId     := 16#0000_0000;   // 信息码回落（R69 点修⑤）：上一轮收割 / 回卷事件不再属当下
                                            // Info codes fall back as a new bypass cycle starts
            bBypassOn    := TRUE;
            uTargetInt   := uInterlockId;
            uSourceInt   := uSourceId;
            WriteLedger(eKind := E_DL_BypassEventKind.eApply);
            eStateInt    := E_DL_BypassState.eBypassed;
        END_IF
        (* 空闲相收到解除沿：无旁路对象，事件不入台账（无中生有即伪造证据） *)
        (* Release edge while idle: nothing to release, not logged *)

    E_DL_BypassState.eBypassed:
        IF fbTrigRel.Q THEN
            (* 本拍解除沿优先于超时迁移（R275）：人工解除即时生效 *)
            (* Release edge outranks the timeout transition in the same scan *)
            bBypassOn  := FALSE;
            uTargetInt := uInterlockId;
            uSourceInt := uSourceId;
            WriteLedger(eKind := E_DL_BypassEventKind.eReleaseByCmd);
            eStateInt  := E_DL_BypassState.eIdle;
        ELSIF tonWindow.Q THEN
            (* 时限到期自动恢复：信息级码（信息级允许每拍重算，本拍一次性落账） *)
            (* Window expired: auto restore, info-level code *)
            bBypassOn  := FALSE;
            uErrorId   := 16#0001_04B1;
            uTargetInt := uInterlockId;
            uSourceInt := uSourceId;
            WriteLedger(eKind := E_DL_BypassEventKind.eReleaseByTimeout);
            eStateInt  := E_DL_BypassState.eIdle;
        END_IF

    E_DL_BypassState.eFault:
        (* 解除路径（R152 自证可达）：复位沿 AND 组态已改对（bWindowInvalid 已消） *)
        (* Clear path: reset edge AND the config is fixed, provably reachable *)
        IF fbTrigReset.Q AND (NOT bWindowInvalid) THEN
            bConfigLatch := FALSE;
            uErrorId     := 16#0000_0000;
            eStateInt    := E_DL_BypassState.eIdle;
        END_IF

    ELSE
        (* 非法状态拦截：不做隐式恢复，直接锁存上报（全库惯用码 0001_0005） *)
        (* Illegal state interception: latch and report, no implicit recovery *)
        eStateInt := E_DL_BypassState.eFault;
        uErrorId  := 16#0001_0005;
        bErrorInt := TRUE;
        bBypassOn := FALSE;      // 迁相补清（R69 点修①）：非法态兜底同样断窗计时 / Same migration clearance

END_CASE;

(*------------------------------------------------------------------------------
 * 段 6｜输出单一出口（范式 P-05）：旁路位只由状态派生一次
 *      Single output exit: the bypass bit derives from the state exactly once
 *      eFault / eIdle 相旁路位必为 FALSE：故障态不携带旁路放行（安全侧）
 *-----------------------------------------------------------------------------*)
bBypassActive  := (eStateInt = E_DL_BypassState.eBypassed);
uBypassCount   := uCntInt;
bLedgerWrapped := (uEventTotal > UDINT#8);
(* 04B2 一次性事件码（R69 点修⑤）：回卷首次发生才发一次，禁每拍重发（信息级可每拍
 * 重算但事件码重发会淹没后续事件码）。回落：复位沿 AND 无组态锁存即归零。 *)
(* Wrap event code is one-shot; it falls back on a reset edge without a config latch *)
IF bLedgerWrapped AND (NOT bWrapCoded) THEN
    uErrorId   := 16#0001_04B2;    // 信息级：台账回卷覆盖 / Info: ledger wrapped
    bWrapCoded := TRUE;            // 一次性标记 / One-shot marker
END_IF
IF fbTrigReset.Q AND (NOT bConfigLatch) THEN
    uErrorId   := 16#0000_0000;    // 信息码随复位沿回落 / Info codes fall back on reset
    bWrapCoded := FALSE;           // 回卷事件码重新武装（再次回卷才重发）/ Re-armed for a later wrap
END_IF
IF UDINT_TO_DINT(uEventTotal) < DINT#8 THEN
    nLedgerCount := DINT_TO_INT(UDINT_TO_DINT(uEventTotal));
ELSE
    nLedgerCount := 8;           // 环形深度即上限 [条] / Ring depth is the cap
END_IF
eLastEvent   := eLastEventInt;
uLastEventSeq := uLastSeqInt;
uLastTarget  := uTargetInt;
uLastSource  := uSourceInt;

FOR nWriteIdx := 0 TO (DL_BYP_RING_DEPTH - 1) DO
    aLedgerKind[nWriteIdx] := aeKindInt[nWriteIdx];     // 台账副本直出 / Ledger copy out
    auLedgerTarget[nWriteIdx] := auiTargetInt[nWriteIdx];
    auLedgerSource[nWriteIdx] := auiSourceInt[nWriteIdx];
END_FOR

bError := bErrorInt OR (eStateInt = E_DL_BypassState.eFault);
eState := eStateInt;
END_FUNCTION_BLOCK

(*------------------------------------------------------------------------------
 * 私有方法: WriteLedger —— 台账环形写入唯一入口（写指针 / 序号 / 计数三记账）
 *      Private method: the single ledger write entry, books pointer, seq and count
 *      调用约定: 仅在本件主体 CASE 内调用；无阻塞、无跨周期状态驻留之外副作用
 *----------------------------------------------------------------------------*)
METHOD WriteLedger
VAR_INPUT
    eKind : E_DL_BypassEventKind;   // 待写事件种类 / Event kind to be written
END_VAR
VAR
    nSlot : INT;                    // 本次写入槽位 [0..7] / Slot index of this write
END_VAR

nSlot := nWriteIdx;                                 // 取当前写指针 / Take the current pointer
aeKindInt[nSlot] := eKind;                          // 事件种类入账 / Kind into the ledger
auiTargetInt[nSlot] := uTargetInt;                  // 目标联锁号入账 / Target id into the ledger
auiSourceInt[nSlot] := uSourceInt;                  // 申请源标识入账 / Source id into the ledger

IF uSeqCounter < DL_BYP_SEQ_MAX THEN
    uSeqCounter := uSeqCounter + 1;                 // 序号推进（饱和）/ Advance sequence, saturating
END_IF
uLastSeqInt   := uSeqCounter;                       // 最近事件序号留影 / Snapshot last sequence
eLastEventInt := eKind;                             // 最近事件种类留影 / Snapshot last kind

IF uCntInt < DL_BYP_CNT_MAX THEN
    uCntInt := uCntInt + 1;                         // 旁路计数推进（255 饱和不回绕）/ Count up, saturating
END_IF

uEventTotal := uEventTotal + 1;                     // 累计事件推进（回卷判据）/ Total events up

nWriteIdx := nWriteIdx + 1;                         // 写指针推进 / Advance the write pointer
IF nWriteIdx >= DL_BYP_RING_DEPTH THEN
    nWriteIdx := 0;                                 // 显式回卷（禁 MOD 方言，IF 等价实现）/ Explicit wrap, IF form
END_IF

END_METHOD

(* ---- FB_DL_RedundantSwitch.st ---- *)
(*==============================================================================
 * 组件名称 (Component)  : FB_DL_RedundantSwitch
 * 所属子库 (Sublibrary) : DL_Base
 * 当前版本 (Version)    : 1.0.0
 * 兼容性   (Platform)   : CODESYS 3.5 / TwinCAT 3 / 汇川 InoProShop / Machine Expert
 *                         仅依赖 Standard.library（TON / R_TRIG / F_TRIG / ABS）
 * 功能描述 (Function)   : 双通道（双传感器或双执行器反馈）冗余选择器。
 *                         持续比较 A/B 偏差，超限并经延时确认后报警；两通道互相矛盾时
 *                         不猜谁对——默认保持最后有效值，也可显式改为跟随某一路或直接判故障；
 *                         单通道失效时按停留时间与速率限制无扰切换到另一通道；
 *                         切换过于频繁则判定抖振并锁存，杜绝"接触器被程序当成振荡器打"。
 *                         解决两个现场通病：①双传感器冗余装了，程序里却只接了一路；
 *                         ②切过去那一瞬间阀门位置跳变，工艺直接甩料。
 *
 * 【核心语义 / Core semantics（边界 B1，本组件最重要的约定）】
 *   两路传感器打架时，程序没有资格替工艺判断谁对。默认策略是 eHoldLast：保持最后
 *   有效值并报警，等工程师到现场看表。要自动跟随某一路，必须显式把 eDevPolicy 改成
 *   eUseA / eUseB，并在设计文件里留档"为什么信这一路"。
 *
 * 【失真与语义披露 / Distortion disclosure】
 *   1) 本块不做 NaN/Inf 检测：IEC 61131-3 无标准判据，各平台行为不一致，强行判断会
 *      引入编译器方言。通道含 NaN 时会污染输出，调用方必须前置量程与断线校验。
 *   2) fMaxSlewRate = 0 的定义是"直接切换"，不是"不切换"。现场若按"0 = 禁用"理解，
 *      会误以为切换失效，故参数注释与手册双重明示。
 *   3) eDevPolicy = eFault 时按"无可用源"口径复用 16#0002_0005：矛盾双方均不可信，
 *      等价于没有可信源。第 4 章未为该策略单列故障码，本块不新造码，改为复用并在此披露。
 *   4) 偏差报警是"已确认事实"，切到单通道后不再有比较对象，因此保持到两路同时有效且
 *      偏差回落，或收到复位沿为止（自检向量 V4）。
 *
 * 开源溯源 (Origin)     : 原创实现（参考西门子 LGF 比较器功能组的公差窗口分类与工业冗余
 *                         惯例的参数域，clean-room 编写，未复制任何源码）
 * 本文件内含       : TYPE  E_DL_RedundancyPriority / E_DL_DeviationPolicy
 *                    TYPE  E_DL_ActiveChannel / E_DL_RedundState
 *                    FB    FB_DL_RedundantSwitch
 * 依赖     (Depends)    : 无 DL_ 内部依赖；Standard.library: TON / R_TRIG / F_TRIG
 * 红线自检 (Redline)    : R1 ✓ 零全局变量表与外部变量引用 ｜ R2 ✓ 零物理 IO 地址直写
 *                         R3 ✓ 纯 IEC 61131-3（无指针、无厂商私有符号）
 *                         R4 ✓ 偏差限钳位 + 时间增量钳位 + 除零前判零 + 抖振锁定
 *                         R5 ✓ 全变量中英双语同行注释 ｜ R6 ✓ 五态 ENUM + CASE + ELSE 兜底
 *                         R7 ✓ 四个实例（一沿 + 三计时）主体最前部无条件刷新
 * 修订历史 (Revision)   :
 *   2026-11-14  v1.0.0  首版入库（Phase 1 收口批次 · R3）
 *============================================================================*)

(*-----------------------------------------------------------------------------
 * 枚举 1: E_DL_RedundancyPriority — 首选通道策略（归属 DL_Base）
 *----------------------------------------------------------------------------*)
TYPE E_DL_RedundancyPriority :
(
    eAuto   := 0,     // 自动：首次选 A，之后跟随当前生效通道 / Auto, pick A first then follow the active one
    eForceA := 1,     // 强制 A，仅在 A 失效时才允许越权到 B / Force A, only A invalidity may override
    eForceB := 2      // 强制 B，仅在 B 失效时才允许越权到 A / Force B, only B invalidity may override
);
END_TYPE

(*-----------------------------------------------------------------------------
 * 枚举 2: E_DL_DeviationPolicy — 偏差超限时的处置策略（归属 DL_Base）
 *----------------------------------------------------------------------------*)
TYPE E_DL_DeviationPolicy :
(
    eHoldLast := 0,   // 保持最后有效值（默认，不猜谁对）/ Hold the last valid value, never guess
    eUseA     := 1,   // 视为 B 漂移，跟随 A / Treat B as drifting, follow A
    eUseB     := 2,   // 视为 A 漂移，跟随 B / Treat A as drifting, follow B
    eFault    := 3    // 偏差超限即判故障（保守工艺）/ Fail on deviation, for conservative processes
);
END_TYPE

(*-----------------------------------------------------------------------------
 * 枚举 3: E_DL_ActiveChannel — 当前生效通道（归属 DL_Base）
 *----------------------------------------------------------------------------*)
TYPE E_DL_ActiveChannel :
(
    eNone := 0,       // 无可用通道 / No usable channel
    eA    := 1,       // 通道 A 生效 / Channel A is active
    eB    := 2        // 通道 B 生效 / Channel B is active
);
END_TYPE

(*-----------------------------------------------------------------------------
 * 枚举 4: E_DL_RedundState — 冗余选择器主状态（归属 DL_Base）
 *----------------------------------------------------------------------------*)
TYPE E_DL_RedundState :
(
    eInit    := 0,    // 初始化（首扫）：按首选策略装载首值 / Initialisation, load the first value per preference
    eNormal  := 10,   // 双通道一致，正常跟随 / Both channels agree, normal tracking
    eSuspect := 20,   // 偏差超限，等待判定 / Deviation confirmed, awaiting a decision
    eRamping := 30,   // 切换过渡中（限速逼近目标）/ Bumpless transition in progress
    eFault   := 99    // 无可用通道或抖振锁定 / No usable channel or chatter latched
);
END_TYPE

(*==============================================================================
 * 功能块: FB_DL_RedundantSwitch
 * 调用约定: 每个扫描周期无条件调用一次，uDeltaTimeMs 必须由调用方注入真实任务间隔。
 *============================================================================*)
FUNCTION_BLOCK FB_DL_RedundantSwitch
VAR_INPUT
    fChannelA       : REAL;                        // 通道 A 测量值 [EU] / Channel A value [EU]
    fChannelB       : REAL;                        // 通道 B 测量值 [EU] / Channel B value [EU]
    bChannelAValid  : BOOL := TRUE;                // A 通道健康（无断线、无超量程）/ A healthy, no wire break
    bChannelBValid  : BOOL := TRUE;                // B 通道健康 / B healthy
    fDeviationLimit : REAL := 1.0;                 // 偏差限 [EU]，合法域 > 0 / Deviation limit [EU], must be > 0
    tDeviationDelay : TIME := T#2S;                // 偏差确认延时 [s]，T#0S = 立即确认 / Confirmation delay [s], T#0S = immediate
    ePreferred      : E_DL_RedundancyPriority := E_DL_RedundancyPriority.eAuto;   // 首选通道策略 / Preferred channel policy
    eDevPolicy      : E_DL_DeviationPolicy := E_DL_DeviationPolicy.eHoldLast;     // 偏差处置策略 / Deviation policy
    tSwitchDwell    : TIME := T#500MS;             // 切换后抑制再次切换的停留时间 [ms] / Post-switch dwell [ms]
    fMaxSlewRate    : REAL := 0.0;                 // 无扰过渡最大变化率 [EU/s]，0 = 直接切换 / Max slew rate, 0 = direct switch
    uDeltaTimeMs    : UDINT;                       // 调用方注入的扫描间隔 [ms] / Injected scan delta [ms]
    fSafeValue      : REAL := 0.0;                 // 双通道失效时的安全值 [EU] / Safe value when no source is usable [EU]
    bReset          : BOOL;                        // 上升沿：复位锁存故障与偏差报警 / Rising edge: reset latched faults
END_VAR
VAR_OUTPUT
    fSelected       : REAL;                        // 选择后的输出值 [EU] / Selected output [EU]
    eActive         : E_DL_ActiveChannel;          // 当前生效通道 / Currently active channel
    bOutputValid    : BOOL;                        // 输出有效（非安全值替代）/ Output valid, not a substituted safe value
    fDeviation      : REAL;                        // 当前偏差 |A-B| [EU]，单通道时恒为 0 / Current deviation, 0 when only one channel
    bDeviationAlarm : BOOL;                        // 偏差报警（已延时确认，保持到回落或复位）/ Deviation alarm, latched until recovery or reset
    bRamping        : BOOL;                        // 过渡进行中 / Bumpless transition in progress
    uSwitchCount    : UDINT;                       // 累计切换次数（饱和）/ Switchover count, saturating
    bError          : BOOL;                        // 故障标志（锁存）/ Fault flag, latched
    uErrorId        : UDINT;                       // 故障码，0 = 无故障 / Error code, 0 = no error
    eState          : E_DL_RedundState;            // 当前状态（供 HMI 诊断）/ Current state for HMI diagnosis
END_VAR
VAR
    fbTrigReset     : R_TRIG;                      // 复位上升沿检测实例 / Reset rising edge detector
    fbTonDev        : TON;                         // 偏差确认定时器 / Deviation confirmation timer
    fbTonDwell      : TON;                         // 切换停留定时器 / Switch dwell timer
    fbTonChatter    : TON;                         // 抖振统计窗口定时器 / Chatter observation window timer
    eStateInt       : E_DL_RedundState;            // 主状态机内部当前态 / Internal state of the main state machine
    eWanted         : E_DL_ActiveChannel;          // 本拍应生效的通道（按策略与有效性推导）/ Channel that should be active this scan
    eTarget         : E_DL_ActiveChannel;          // 过渡目标通道 / Ramp target channel
    ePending        : E_DL_ActiveChannel;          // 本拍待发起的切换目标，eNone = 无 / Pending switch target, eNone = none
    fSelectedInt    : REAL;                        // 输出值内部副本（单一出口用）/ Internal copy of the output, for the single exit
    fTargetVal      : REAL;                        // 过渡目标值 [EU] / Ramp target value [EU]
    fLastValid      : REAL;                        // 最后有效值 [EU]，保持策略的锚点 / Last valid value, the anchor of the hold policy
    fStep           : REAL;                        // 本拍允许的最大变化量 [EU] / Maximum allowed change this scan [EU]
    fDevLimEff      : REAL;                        // 钳位后的偏差限 [EU] / Clamped deviation limit [EU]
    fDtSec          : REAL;                        // 扫描间隔换算成秒 [s] / Scan delta in seconds [s]
    tDwellEff       : TIME;                        // 钳位后的停留时间 [ms] / Clamped dwell time [ms]
    uDtEff          : UDINT;                       // 钳位后的扫描间隔 [ms] / Clamped scan delta [ms]
    uSwInt          : UDINT;                       // 切换次数内部副本（饱和）/ Internal switch counter, saturating
    uWarnId         : UDINT;                       // 本拍瞬时告警码（不进锁存）/ Instantaneous warning code of this scan
    nChatterCnt     : INT;                         // 统计窗口内的切换计数 / Switch count inside the observation window
    bDwellRun       : BOOL;                        // 停留计时进行中（TRUE = 禁止再切）/ Dwell timer running, switching inhibited
    bAnyValid       : BOOL;                        // 至少一路有效 / At least one channel is valid
    bBothValid      : BOOL;                        // 两路同时有效 / Both channels are valid
    bActiveValid    : BOOL;                        // 当前生效通道仍然有效 / The active channel is still valid
    bTargetValid    : BOOL;                        // 过渡目标通道仍然有效 / The ramp target is still valid
    bSwitchNeed     : BOOL;                        // 本拍需要切换（已含停留抑制）/ Switching required this scan
    bAlarmInt       : BOOL;                        // 偏差报警内部副本 / Internal copy of the deviation alarm
    bChatterTrip    : BOOL;                        // 抖振判据成立 / Chatter criterion satisfied
    bFirstScan      : BOOL := TRUE;                // 上电首扫标志 / First-scan flag
END_VAR
VAR CONSTANT
    DL_RS_DEV_MIN     : REAL := 1.0E-6;            // 偏差限下限 [EU]，兼作浮点判零容差 / Deviation-limit floor, doubles as epsilon
    DL_RS_CHATTER_MAX : INT  := 5;                 // 窗口内允许的最大切换次数 / Max switches per observation window
    DL_RS_CHATTER_WIN : TIME := T#10S;             // 抖振统计窗口 [s] / Chatter observation window [s]
    DL_RS_DT_MAX      : UDINT := 60000;            // 时间增量上限 [ms]，防长时间断点造成巨跳 / Delta clamp [ms]
    DL_RS_CNT_MAX     : UDINT := 16#FFFF_FFFE;     // 切换计数器饱和值 / Switch counter saturation
    DL_RS_DWELL_MAX   : TIME := T#1H;              // 停留时间上限钳位 [s] / Dwell upper clamp [s]
    DL_RS_MS_PER_S    : REAL := 1000.0;            // 毫秒换算常数 [ms/s] / Milliseconds per second
END_VAR

(*------------------------------------------------------------------------------
 * 段 1｜无条件刷新区（红线 R7）：一沿 + 三计时器，全部位于主体最前部
 *      Unconditional refresh zone: one edge and three timers at the very top
 *      定时器 IN 先由"原始输入 + 上一拍参数"推导成 BOOL，实例调用本身绝不进 IF
 *      偏差限取自上一拍的钳位值，滞后一拍对"确认延时"这种秒级量无影响
 *-----------------------------------------------------------------------------*)
fbTrigReset(CLK := bReset);

(* 停留时间钳位先于计时器：超长停留会让人误以为切换失效，钳到 1 h 并保持可观测 *)
(* Clamp the dwell before the timer call so the timer never gets an absurd PT *)
IF tSwitchDwell > DL_RS_DWELL_MAX THEN
    tDwellEff := DL_RS_DWELL_MAX;
ELSE
    tDwellEff := tSwitchDwell;
END_IF

fbTonDev(IN := bChannelAValid AND bChannelBValid AND (ABS(fChannelA - fChannelB) > fDevLimEff),
         PT := tDeviationDelay);

fbTonDwell(IN := bDwellRun, PT := tDwellEff);

fbTonChatter(IN := (nChatterCnt > 0), PT := DL_RS_CHATTER_WIN);

IF fbTonDwell.Q THEN
    bDwellRun := FALSE;
END_IF

IF fbTonChatter.Q THEN
    nChatterCnt := 0;
END_IF

(*------------------------------------------------------------------------------
 * 段 2｜上电首扫：状态、通道号与输出必须显式落到安全侧，不能依赖默认零
 *      First-scan init: state, channel and output are forced to the safe side
 *-----------------------------------------------------------------------------*)
IF bFirstScan THEN
    bFirstScan   := FALSE;
    eStateInt    := E_DL_RedundState.eInit;
    eActive      := E_DL_ActiveChannel.eNone;
    eTarget      := E_DL_ActiveChannel.eNone;
    ePending     := E_DL_ActiveChannel.eNone;
    fSelectedInt := fSafeValue;
    fLastValid   := fSafeValue;
    nChatterCnt  := 0;
    bDwellRun    := FALSE;
END_IF

(*------------------------------------------------------------------------------
 * 段 2b｜故障码口径（红线 R15）：锁存期保留进入故障时的码，瞬时告警不得覆盖它
 *      Error-code policy: instantaneous warnings must never overwrite a latched code
 *      先把瞬时码收进 uWarnId，等确认当前不在故障锁存里才落到 uErrorId
 *-----------------------------------------------------------------------------*)
uWarnId := 16#0000;

(*------------------------------------------------------------------------------
 * 段 3｜时间增量校验（边界 B3/B8）：0 或超上限一律钳位并告警
 *      Delta-time check: zero or over-limit values are clamped and reported
 *      0 会让过渡停走（每拍增量 0）；回绕值会把运行方向算反，都不可接受
 *-----------------------------------------------------------------------------*)
IF uDeltaTimeMs = 0 THEN
    uDtEff   := 1;
    uWarnId  := 16#0001_0008;
ELSIF uDeltaTimeMs > DL_RS_DT_MAX THEN
    uDtEff   := DL_RS_DT_MAX;
    uWarnId  := 16#0001_0008;
ELSE
    uDtEff := uDeltaTimeMs;
END_IF

fDtSec := UDINT_TO_REAL(uDtEff) / DL_RS_MS_PER_S;

(*------------------------------------------------------------------------------
 * 段 4｜偏差限钳位（边界 B7）：先取绝对值再钳下限，负号视为"填错符号"
 *      Deviation-limit clamp: absolute value first, then floor at the epsilon
 *      偏差限为 0 会让任何微小噪声都报警，必须抬到 1E-6 而不是放行
 *-----------------------------------------------------------------------------*)
fDevLimEff := ABS(fDeviationLimit);

IF fDevLimEff < DL_RS_DEV_MIN THEN
    fDevLimEff := DL_RS_DEV_MIN;
    uWarnId    := 16#0001_0001;
END_IF

(* 瞬时告警落码：故障锁存期间一律不落码，保证 HMI 读到的根因不被参数告警冲掉 *)
(* Warnings land only outside the latched fault state, otherwise the root cause is lost *)
IF eStateInt <> E_DL_RedundState.eFault THEN
    IF uWarnId <> 16#0000 THEN
        uErrorId := uWarnId;
    ELSE
        uErrorId := 16#0000_0000;
    END_IF
END_IF

(*------------------------------------------------------------------------------
 * 段 5｜有效性与偏差（边界 B6 的前置量）：单通道时偏差恒为 0
 *      Validity and deviation: with one channel there is no comparison object
 *      单通道时"沿用旧偏差"会让报警永远挂着，必须显式归零
 *-----------------------------------------------------------------------------*)
bAnyValid  := bChannelAValid OR bChannelBValid;
bBothValid := bChannelAValid AND bChannelBValid;

IF bBothValid THEN
    fDeviation := ABS(fChannelA - fChannelB);
ELSE
    fDeviation := 0.0;
END_IF

(*------------------------------------------------------------------------------
 * 段 6｜偏差报警（边界：V4 语义）：确认后保持，回落或复位才清
 *      Deviation alarm: latched once confirmed, cleared on recovery or reset
 *-----------------------------------------------------------------------------*)
IF fbTonDev.Q THEN
    bAlarmInt := TRUE;
END_IF

IF bBothValid AND (fDeviation <= fDevLimEff) THEN
    bAlarmInt := FALSE;
END_IF

IF fbTrigReset.Q THEN
    bAlarmInt := FALSE;
END_IF

(*------------------------------------------------------------------------------
 * 段 7｜目标通道推导（边界 B1/B2）
 *      Target-channel derivation: preference first, then validity, never both guesses
 *      eAuto 的语义是"保持当前有效通道"，只有当前通道失效才换——不是每拍重新投票
 *-----------------------------------------------------------------------------*)
IF NOT bAnyValid THEN
    eWanted := E_DL_ActiveChannel.eNone;
ELSIF ePreferred = E_DL_RedundancyPriority.eForceA THEN
    IF bChannelAValid THEN
        eWanted := E_DL_ActiveChannel.eA;
    ELSE
        eWanted := E_DL_ActiveChannel.eB;
    END_IF
ELSIF ePreferred = E_DL_RedundancyPriority.eForceB THEN
    IF bChannelBValid THEN
        eWanted := E_DL_ActiveChannel.eB;
    ELSE
        eWanted := E_DL_ActiveChannel.eA;
    END_IF
ELSE
    (* eAuto：当前通道仍有效就不动，失效才换到另一路 *)
    IF (eActive = E_DL_ActiveChannel.eA) AND bChannelAValid THEN
        eWanted := E_DL_ActiveChannel.eA;
    ELSIF (eActive = E_DL_ActiveChannel.eB) AND bChannelBValid THEN
        eWanted := E_DL_ActiveChannel.eB;
    ELSIF bChannelAValid THEN
        eWanted := E_DL_ActiveChannel.eA;
    ELSE
        eWanted := E_DL_ActiveChannel.eB;
    END_IF
END_IF

(*------------------------------------------------------------------------------
 * 段 8｜切换判据（边界 B5）：源通道失效可越权（安全优先），否则受停留时间抑制
 *      Switch criterion: a dead source overrides the dwell, a healthy one does not
 *-----------------------------------------------------------------------------*)
IF eActive = E_DL_ActiveChannel.eA THEN
    bActiveValid := bChannelAValid;
ELSIF eActive = E_DL_ActiveChannel.eB THEN
    bActiveValid := bChannelBValid;
ELSE
    bActiveValid := FALSE;
END_IF

bSwitchNeed := (eWanted <> E_DL_ActiveChannel.eNone)
               AND (eWanted <> eActive)
               AND ((NOT bDwellRun) OR (NOT bActiveValid));

(*------------------------------------------------------------------------------
 * 段 9｜主状态机（红线 R6）：ENUM + CASE + ELSE 兜底
 *      Main state machine with the mandatory ELSE fallback
 *-----------------------------------------------------------------------------*)
ePending := E_DL_ActiveChannel.eNone;

CASE eStateInt OF

    E_DL_RedundState.eInit:
        (* 首扫后按策略装载首值；双无效直接进故障，输出安全值 *)
        (* Load the first value per preference; no valid source goes straight to fault *)
        IF bAnyValid THEN
            eActive      := eWanted;
            IF eActive = E_DL_ActiveChannel.eA THEN
                fSelectedInt := fChannelA;
            ELSE
                fSelectedInt := fChannelB;
            END_IF
            fLastValid := fSelectedInt;
            eTarget    := eActive;
            fTargetVal := fSelectedInt;
            eStateInt  := E_DL_RedundState.eNormal;
        ELSE
            eStateInt := E_DL_RedundState.eFault;
            uErrorId  := 16#0002_0005;
        END_IF

    E_DL_RedundState.eNormal:
        IF NOT bAnyValid THEN
            eStateInt := E_DL_RedundState.eFault;
            uErrorId  := 16#0002_0005;
        ELSIF bSwitchNeed THEN
            ePending  := eWanted;
            eStateInt := E_DL_RedundState.eRamping;
        ELSIF fbTonDev.Q THEN
            (* 偏差确认到期：进入疑似态，由策略决定输出与后续动作 *)
            (* Deviation confirmed: enter the suspect state, the policy decides *)
            eStateInt := E_DL_RedundState.eSuspect;
        ELSE
            (* 正常跟随：输出必须每拍跟踪当前生效通道，否则会输出一个冻结值 *)
            (* Normal tracking: the output must follow the active channel every scan *)
            IF (eActive = E_DL_ActiveChannel.eA) AND bChannelAValid THEN
                fSelectedInt := fChannelA;
            ELSIF (eActive = E_DL_ActiveChannel.eB) AND bChannelBValid THEN
                fSelectedInt := fChannelB;
            END_IF
            fLastValid := fSelectedInt;
        END_IF

    E_DL_RedundState.eSuspect:
        IF NOT bAnyValid THEN
            eStateInt := E_DL_RedundState.eFault;
            uErrorId  := 16#0002_0005;
        ELSIF bSwitchNeed THEN
            (* 疑似失效的那一路被宣告 Valid = FALSE：偏差比较已无意义，直接切 *)
            (* The suspect channel dropped its valid flag: compare is meaningless, switch at once *)
            ePending  := eWanted;
            eStateInt := E_DL_RedundState.eRamping;
        ELSIF (NOT bBothValid) OR (fDeviation <= fDevLimEff) THEN
            (* 偏差已无对象或已回落：回到正常跟随 *)
            (* No comparison object left, or the deviation recovered: back to normal *)
            eStateInt := E_DL_RedundState.eNormal;
        ELSE
            CASE eDevPolicy OF
                E_DL_DeviationPolicy.eHoldLast:
                    (* 默认：保持最后有效值，谁都不信 *)
                    (* Default: hold the last valid value, trust neither channel *)
                    fSelectedInt := fLastValid;

                E_DL_DeviationPolicy.eUseA:
                    IF bChannelAValid THEN
                        fSelectedInt := fChannelA;
                        fLastValid   := fSelectedInt;
                    ELSE
                        fSelectedInt := fLastValid;
                    END_IF

                E_DL_DeviationPolicy.eUseB:
                    IF bChannelBValid THEN
                        fSelectedInt := fChannelB;
                        fLastValid   := fSelectedInt;
                    ELSE
                        fSelectedInt := fLastValid;
                    END_IF

                E_DL_DeviationPolicy.eFault:
                    (* 保守工艺：矛盾即停机，按"无可用源"口径复用 0002_0005（见头注释） *)
                    (* Conservative: contradictory means stop, reuse 0002_0005 as documented *)
                    eStateInt := E_DL_RedundState.eFault;
                    uErrorId  := 16#0002_0005;

                ELSE
                    eStateInt := E_DL_RedundState.eFault;
                    uErrorId  := 16#0001_0005;
            END_CASE
        END_IF

    E_DL_RedundState.eRamping:
        IF eTarget = E_DL_ActiveChannel.eA THEN
            bTargetValid := bChannelAValid;
        ELSIF eTarget = E_DL_ActiveChannel.eB THEN
            bTargetValid := bChannelBValid;
        ELSE
            bTargetValid := FALSE;
        END_IF

        (* 目标通道的物理值在过渡期间仍会变，目标值必须每拍刷新，否则会爬向一个陈旧值 *)
        (* The target channel keeps moving during the ramp, so refresh the target value each scan *)
        IF bTargetValid THEN
            IF eTarget = E_DL_ActiveChannel.eA THEN
                fTargetVal := fChannelA;
            ELSE
                fTargetVal := fChannelB;
            END_IF
        END_IF

        IF NOT bAnyValid THEN
            eStateInt := E_DL_RedundState.eFault;
            uErrorId  := 16#0002_0005;
        ELSIF NOT bTargetValid THEN
            (* 目标在过渡途中失效：中止过渡，退回当前生效通道，不产生第二次切换计数 *)
            (* Target died mid-ramp: abort and retreat, without counting a second switch *)
            eTarget    := eActive;
            fTargetVal := fSelectedInt;
            eStateInt  := E_DL_RedundState.eNormal;
        ELSIF (ABS(fMaxSlewRate) <= DL_RS_DEV_MIN) OR (fDtSec <= 0.0) THEN
            (* 边界 B4：速率 0 定义为直接切换；dt 异常时也取向直接吸附，绝不发散的慢慢爬 *)
            (* Rate 0 means direct switching; an abnormal dt snaps instead of crawling forever *)
            fSelectedInt := fTargetVal;
            eActive      := eTarget;
            fLastValid   := fSelectedInt;
            eStateInt    := E_DL_RedundState.eNormal;
        ELSE
            fStep := ABS(fMaxSlewRate) * fDtSec;
            IF ABS(fTargetVal - fSelectedInt) <= fStep THEN
                fSelectedInt := fTargetVal;
                eActive      := eTarget;
                fLastValid   := fSelectedInt;
                eStateInt    := E_DL_RedundState.eNormal;
            ELSE
                IF fTargetVal > fSelectedInt THEN
                    fSelectedInt := fSelectedInt + fStep;
                ELSE
                    fSelectedInt := fSelectedInt - fStep;
                END_IF
            END_IF
        END_IF

    E_DL_RedundState.eFault:
        (* 边界 B6：双通道失效时输出安全值，绝不输出"最后有效值"——最后值同样可疑 *)
        (* Both channels dead: output the safe value, never the last valid one *)
        fSelectedInt := fSafeValue;
        IF fbTrigReset.Q AND bAnyValid THEN
            uErrorId    := 16#0000_0000;
            nChatterCnt := 0;
            bDwellRun   := FALSE;
            eStateInt   := E_DL_RedundState.eInit;
        END_IF

    ELSE
        (* 非法状态拦截：不做隐式恢复，直接锁存上报 *)
        (* Illegal state interception: no implicit recovery, latch and report *)
        eStateInt := E_DL_RedundState.eFault;
        uErrorId  := 16#0001_0005;

END_CASE;

(*------------------------------------------------------------------------------
 * 段 10｜切换提交（唯一切换记账点）
 *      Switch commitment: the one and only place where switching is booked
 *      只在状态机确实发起切换的那一拍记账，过渡期内绝不重复累加，否则抖振判据必被误触
 *      Bookkeeping happens once per initiated switch, never during the ramp itself
 *-----------------------------------------------------------------------------*)
IF ePending <> E_DL_ActiveChannel.eNone THEN

    eTarget := ePending;

    IF eTarget = E_DL_ActiveChannel.eA THEN
        fTargetVal := fChannelA;
    ELSE
        fTargetVal := fChannelB;
    END_IF

    IF uSwInt < DL_RS_CNT_MAX THEN
        uSwInt := uSwInt + 1;
    ELSE
        uErrorId := 16#0001_0007;
    END_IF

    (* 计数封顶在 MAX+1，既能判定越限又不会让 INT 溢出 *)
    (* The counter stops at MAX+1: enough to trip, never enough to overflow *)
    IF nChatterCnt <= DL_RS_CHATTER_MAX THEN
        nChatterCnt := nChatterCnt + 1;
    END_IF

    bDwellRun := TRUE;

    (* 抖振判据（边界 B6）：窗口内切换次数超限即锁定，说明设定错误或信号在临界点抖 *)
    (* Chatter: too many switches inside the window means a bad setup or a dithering signal *)
    bChatterTrip := (nChatterCnt > DL_RS_CHATTER_MAX);
    IF bChatterTrip THEN
        uErrorId  := 16#0002_0006;
        eStateInt := E_DL_RedundState.eFault;
    ELSE
        (* 边界 B4：速率 0 定义为"直接切换"，在发起的同一拍吸附到目标值 *)
        (* Rate 0 means a direct switch: snap to the target in the very same scan *)
        IF ABS(fMaxSlewRate) <= DL_RS_DEV_MIN THEN
            fSelectedInt := fTargetVal;
            eActive      := eTarget;
            fLastValid   := fSelectedInt;
            eStateInt    := E_DL_RedundState.eNormal;
        END_IF
    END_IF

END_IF

(*------------------------------------------------------------------------------
 * 段 11｜输出单一出口（范式 P-05）
 *      Single output exit: every output is derived once, here
 *-----------------------------------------------------------------------------*)
fSelected       := fSelectedInt;
bOutputValid    := bAnyValid AND (eActive <> E_DL_ActiveChannel.eNone)
                   AND (eStateInt <> E_DL_RedundState.eFault);
bDeviationAlarm := bAlarmInt;
bRamping        := (eStateInt = E_DL_RedundState.eRamping);
uSwitchCount    := uSwInt;
bError          := (eStateInt = E_DL_RedundState.eFault);
eState          := eStateInt;
END_FUNCTION_BLOCK

(* ---- FC_DL_BitRotateEx.st ---- *)
//==============================================================================
// 函数：FC_DL_BitRotateEx ｜ 中文名称：位串循环移位（跨位回卷）
// 所属子库：DL_Base ｜ 版本：v1.0.0 ｜ 日期：2026-11-23
// 兼容：CODESYS V3.5+ / TwinCAT 3 / 汇川 InoProShop（纯标准库 SHL/SHR 组合）
// 功能描述：位串循环移位原子：左/右方向 × 8/16/32 位宽度域内回卷。
//           实现口径：SHL(x,n) OR SHR(x,w−n) 组合回卷，n 先归一到
//           [0, w−1]（负移位量取模回卷，禁 SHL(x,位宽) 未定义行为——
//           移位量归一后为 0 时直通返回原值，落位组合分支的移位量恒在
//           1..w−1 安全域）。与 ShlEx/ShrEx 邻件分工：那两件做饱和/截断
//           单向移位，本件只做回卷循环移位，互不替代。
// 开源溯源 (Origin)：原创实现（t0-std-wrapper 包装族补口，零外部源码行，
//           clean-room 独立编写；与 ShlEx/ShrEx 邻件分工已在头注释声明）
// 公开接口清单：输入 dwVal / nShift / eDir / eWidth；输出 dwRotated / bValid
// 错误码表：纯函数无状态机码轨；无效输入经 bValid = FALSE 表达（哨兵返回
//           0.0），本件不占用 16#0001 段码位（邻件免让位）
// 状态机：E_DL_RotDir / E_DL_RotWidth（本文件唯一定义，全库唯一属主）：
//           方向 eLeft = 0 / eRight = 1；宽度 eW8 = 8 / eW16 = 16 / eW32 = 32
// 边界行为：① 移位量任意整数（含负值）先 MOD 归一到 [0, w−1]；
//           ② 归一后为 0 直通返回原值（组合分支移位量恒 1..w−1，禁
//             SHL(x,位宽) 未定义行为）；
//           ③ 宽度域外（非 8/16/32）→ 哨兵 0.0 返回；
//           ④ 回卷结果按宽度掩码截取（高位残留清零）。
// 修订历史：v1.0.0 2026-11-23 首版（R73 派单 · 批 3 · 序 12）
//==============================================================================

(*------------------------------------------------------------------------------
 * 枚举: E_DL_RotDir / E_DL_RotWidth（归属本函数，同文件发布，全库唯一属主）
 * 含义: 移位方向与位串宽度域，成员与 CASE 标签双向完备。
 *-----------------------------------------------------------------------------*)
TYPE E_DL_RotDir :
(
    eLeft  := 0,   // 左循环移位 / Rotate left
    eRight := 1    // 右循环移位 / Rotate right
);
END_TYPE

TYPE E_DL_RotWidth :
(
    eW8  := 8,     // 8 位宽度域 / 8-bit width domain
    eW16 := 16,    // 16 位宽度域 / 16-bit width domain
    eW32 := 32     // 32 位宽度域 / 32-bit width domain
);
END_TYPE

(*------------------------------------------------------------------------------
 * 调用示例：dwR := FC_DL_BitRotateEx(dwVal := 16#0000_00A1,
 *             nShift := 3, eDir := E_DL_RotDir.eLeft,
 *             eWidth := E_DL_RotWidth.eW8, bValid => bOk);
 * 注意：移位量先归一回卷，任意整数（含负）均合法；宽度域外拒绝。
 *-----------------------------------------------------------------------------*)
FUNCTION FC_DL_BitRotateEx : DWORD
VAR_INPUT
    dwVal   : DWORD;                   // 输入位串 [—] / Input bit pattern
    nShift  : DINT;                    // 移位量 [位]，任意整数（含负，取模回卷）/ Shift amount [bits], any integer, wrapped by modulo
    eDir    : E_DL_RotDir;             // 移位方向枚举 [—] / Rotation direction enum
    eWidth  : E_DL_RotWidth;           // 位串宽度域枚举 [位] / Width domain enum [bits]
END_VAR
VAR_OUTPUT
    bValid  : BOOL;                    // 结果有效标志，FALSE 时返回哨兵 0.0 / Result validity flag
END_VAR
VAR
    nW      : DINT;                    // 生效宽度 [位] / Effective width [bits]
    nEff    : DINT;                    // 归一后移位量 [位]，域 0..w−1 / Normalized shift [bits], range 0..w-1
    dwMask  : DWORD;                   // 宽度掩码 / Width mask
    dwLo    : DWORD;                   // 回卷低位段 / Wrapped low segment
    dwHi    : DWORD;                   // 回卷高位段 / Wrapped high segment
END_VAR
VAR CONSTANT
    DW_ROT_SENTINEL : DWORD := 16#0000_0000; // 无效哨兵返回值 / Sentinel return for invalid
END_VAR

// ---- 段 1｜出口默认值（纯函数无实例，无定时器/沿刷新义务）----
bValid := FALSE;                      // 缺省无效 / Invalid by default

// ---- 段 2｜宽度域解析（CASE 带 ELSE；非法宽度拒绝）----
CASE eWidth OF
    E_DL_RotWidth.eW8:                 // 8 位域：掩码低 8 位 / 8-bit domain
        nW     := 8;                   // 生效宽度 [位] / Effective width
        dwMask := 16#0000_00FF;        // 宽度掩码 / Width mask
    E_DL_RotWidth.eW16:                // 16 位域：掩码低 16 位 / 16-bit domain
        nW     := 16;                  // 生效宽度 [位] / Effective width
        dwMask := 16#0000_FFFF;        // 宽度掩码 / Width mask
    E_DL_RotWidth.eW32:                // 32 位域：全掩码 / 32-bit domain
        nW     := 32;                  // 生效宽度 [位] / Effective width
        dwMask := 16#FFFF_FFFF;        // 宽度掩码 / Width mask
    ELSE                               // 枚举非法值兜底（R21：CASE 必带 ELSE）
        FC_DL_BitRotateEx := DW_ROT_SENTINEL; // 非法宽度：哨兵零返回 / Illegal width, sentinel zero return
        RETURN;                        // 结构早退 / early exit
END_CASE

// ---- 段 3｜移位量归一：MOD 取模 + 双侧回卷（负移位量合法）----
nEff := nShift MOD nW;                // 先取模（可能为负，DINT MOD 语义随被除数）/ Modulo first, may be negative
IF nEff < 0 THEN
    nEff := nEff + nW;                // 负移位量回卷到 [0, w−1] / Negative shift wrapped up
END_IF

// ---- 段 4｜回卷主体：移位量 0 直通；组合分支移位量恒 1..w−1 安全域 ----
IF nEff = 0 THEN
    FC_DL_BitRotateEx := dwVal AND dwMask; // 零移位直通（掩码截取）/ Zero shift pass-through, masked
ELSE
    IF eDir = E_DL_RotDir.eLeft THEN  // 左循环：高段出环回低位
        dwHi := SHL(dwVal AND dwMask, DINT_TO_UINT(nEff));        // 左移高位段（标准显式转换 R10）/ Left-shifted high segment, standard explicit cast
        dwLo := SHR(dwVal AND dwMask, DINT_TO_UINT(nW - nEff));   // 出环段回卷到低位 / Wrapped-out segment to low bits
        FC_DL_BitRotateEx := (dwHi OR dwLo) AND dwMask; // 回卷合成 + 掩码截取 / Rotated blend, masked
    ELSE                              // 右循环（含枚举非法值并入右旋，方向枚举仅两员）
        dwLo := SHR(dwVal AND dwMask, DINT_TO_UINT(nEff));        // 右移低位段 / Right-shifted low segment
        dwHi := SHL(dwVal AND dwMask, DINT_TO_UINT(nW - nEff));   // 出环段回卷到高位 / Wrapped-out segment to high bits
        FC_DL_BitRotateEx := (dwHi OR dwLo) AND dwMask; // 回卷合成 + 掩码截取 / Rotated blend, masked
    END_IF
END_IF
bValid := TRUE;                       // 全部防御通过：结果有效 / Result valid
END_FUNCTION

(* ---- FC_DL_ConcUnitConvert.st ---- *)
(*
  FC_DL_ConcUnitConvert —— 浓度换算 ppm 与 % 与 mg/L
  分类：DL_Base | 复杂度：1 | 轮次：R86
  开源溯源：道莅原创（clean-room 自研，纯 IEC 61131-3 通用算法），无外部代码引用
  许可证：MIT
  职责：把三种浓度单位统一折算到基准单位 mg/L（稀溶液口径：1 ppm ≈ 1 mg/L；1 % = 10000 mg/L）。
  契约：fIn 输入值 [源单位]，eUnit 源单位枚举；fOut 折算结果 [mg/L]；返回 TRUE 表示 fOut 可信。
  边界：① 稀溶液近似已显式声明，高浓度 / 非水基介质不得直接套用；② 未知枚举 / 非有限输入 → FALSE + 0.0 哨兵；
        ③ 无除法，零全局、零物理地址、零库件依赖。
*)

(*-----------------------------------------------------------------------------
 * 枚举: E_DL_CncUnit（浓度单位，归属本文件，全库唯一定义）
 *----------------------------------------------------------------------------*)
TYPE E_DL_CncUnit :
(
    eMgPerL   := 0,    // 毫克每升（基准单位，稀溶液近似等于 ppm） [mg/L] / Milligram per litre, the base unit
    ePpm      := 1,    // 百万分之一（体积比，稀溶液按 1 mg/L 折算） [ppm] / Parts per million, approximated
    ePercent  := 2     // 百分比浓度（= 10000 mg/L） [%] / Percent concentration
);
END_TYPE

FUNCTION FC_DL_ConcUnitConvert : BOOL
VAR_INPUT
    fIn   : LREAL := 0.0;              // 输入值 [源单位] / The input value in the source unit
    eUnit : E_DL_CncUnit;              // 源单位枚举 [—] / The source unit enumeration
END_VAR
VAR_OUTPUT
    fOut : LREAL;                      // 折算结果 [mg/L] / The converted value in the base unit
END_VAR
VAR CONSTANT
    DL_CN_PPM : LREAL := 1.0;          // 1 ppm 折 mg/L 的系数（稀溶液） [-] / ppm to mg per litre, dilute solution
    DL_CN_PCT : LREAL := 10000.0;      // 1 % 折 mg/L 的系数 [-] / percent to mg per litre
    DL_CN_INF : LREAL := 1.0E30;       // 非有限 / 越界判据上限 [-] / The magnitude gate
    DL_CN_Z   : LREAL := 0.0;          // 浮点零常量 [mg/L] / The floating point zero constant
END_VAR

FC_DL_ConcUnitConvert := FALSE;                           // 返回值预置假 / preset the return false
fOut := DL_CN_Z;                                          // 输出预置零哨兵 [mg/L] / preset the zero sentinel
IF (fIn <> fIn) OR (ABS(fIn) > DL_CN_INF) THEN            // 自反判 NaN 或越限判 Inf / NaN or Inf
    fOut := DL_CN_Z;                                      // 非有限值输出零哨兵 [mg/L] / zero the non finite input
ELSE
    CASE eUnit OF
        E_DL_CncUnit.eMgPerL:                             // 基准单位直通 / the base unit passes through
            fOut := fIn;                                  // 直通不换算 [mg/L] / pass through unchanged
            FC_DL_ConcUnitConvert := TRUE;                // 结果可信 / the result is valid
        E_DL_CncUnit.ePpm:                                // 百万分之一（体积比） / parts per million
            fOut := fIn * DL_CN_PPM;                      // 按稀溶液 1:1 折算 [mg/L] / dilute solution conversion
            FC_DL_ConcUnitConvert := TRUE;                // 结果可信 / the result is valid
        E_DL_CncUnit.ePercent:                            // 百分比浓度 / percent concentration
            fOut := fIn * DL_CN_PCT;                      // 乘 10000 [mg/L] / multiply by the factor
            FC_DL_ConcUnitConvert := TRUE;                // 结果可信 / the result is valid
    ELSE
        fOut := DL_CN_Z;                                  // 未知枚举输出零哨兵 [mg/L] / zero sentinel on an unknown unit
        FC_DL_ConcUnitConvert := FALSE;                   // 未知枚举不可信 / an unknown unit is not valid
    END_CASE
END_IF
END_FUNCTION

(* ---- FC_DL_CurrentUnitConvert.st ---- *)
(*
  FC_DL_CurrentUnitConvert —— 电流换算 A/mA/kA
  分类：DL_Base | 复杂度：1 | 轮次：R86
  开源溯源：道莅原创（clean-room 自研，纯 IEC 61131-3 通用算法），无外部代码引用
  许可证：MIT
  职责：把电流统一折算到基准单位 A：A 直通、mA 乘 0.001、kA 乘 1000。
  契约：fIn 输入值 [源单位]，eUnit 源单位枚举；fOut 折算结果 [A]；返回 TRUE 表示 fOut 可信。
  边界：未知枚举 / 非有限输入 → 返回 FALSE，fOut 给 0.0 哨兵；无除法，零全局、零物理地址、零库件依赖。
*)

(*-----------------------------------------------------------------------------
 * 枚举: E_DL_CurUnit（电流单位，归属本文件，全库唯一定义）
 *----------------------------------------------------------------------------*)
TYPE E_DL_CurUnit :
(
    eAmpere   := 0,    // 安培（基准单位） [A] / Ampere, the base unit
    eMilliAmp := 1,    // 毫安 [mA] / Milliampere
    eKiloAmp  := 2     // 千安 [kA] / Kiloampere
);
END_TYPE

FUNCTION FC_DL_CurrentUnitConvert : BOOL
VAR_INPUT
    fIn   : LREAL := 0.0;              // 输入值 [源单位] / The input value in the source unit
    eUnit : E_DL_CurUnit;              // 源单位枚举 [—] / The source unit enumeration
END_VAR
VAR_OUTPUT
    fOut : LREAL;                      // 折算结果 [A] / The converted value in the base unit
END_VAR
VAR CONSTANT
    DL_CU_MA  : LREAL := 0.001;        // 1 mA 折 A 的系数 [-] / milliampere to ampere
    DL_CU_KA  : LREAL := 1000.0;       // 1 kA 折 A 的系数 [-] / kiloampere to ampere
    DL_CU_INF : LREAL := 1.0E30;       // 非有限 / 越界判据上限 [-] / The magnitude gate
    DL_CU_Z   : LREAL := 0.0;          // 浮点零常量 [A] / The floating point zero constant
END_VAR

FC_DL_CurrentUnitConvert := FALSE;                        // 返回值预置假 / preset the return false
fOut := DL_CU_Z;                                          // 输出预置零哨兵 [A] / preset the zero sentinel
IF (fIn <> fIn) OR (ABS(fIn) > DL_CU_INF) THEN            // 自反判 NaN 或越限判 Inf / NaN or Inf
    fOut := DL_CU_Z;                                      // 非有限值输出零哨兵 [A] / zero the non finite input
ELSE
    CASE eUnit OF
        E_DL_CurUnit.eAmpere:                             // 基准单位直通 / the base unit passes through
            fOut := fIn;                                  // 直通不换算 [A] / pass through unchanged
            FC_DL_CurrentUnitConvert := TRUE;             // 结果可信 / the result is valid
        E_DL_CurUnit.eMilliAmp:                           // 毫安折安 / milliampere to ampere
            fOut := fIn * DL_CU_MA;                       // 乘 0.001 [A] / multiply by the factor
            FC_DL_CurrentUnitConvert := TRUE;             // 结果可信 / the result is valid
        E_DL_CurUnit.eKiloAmp:                            // 千安折安 / kiloampere to ampere
            fOut := fIn * DL_CU_KA;                       // 乘 1000 [A] / multiply by the factor
            FC_DL_CurrentUnitConvert := TRUE;             // 结果可信 / the result is valid
    ELSE
        fOut := DL_CU_Z;                                  // 未知枚举输出零哨兵 [A] / zero sentinel on an unknown unit
        FC_DL_CurrentUnitConvert := FALSE;                // 未知枚举不可信 / an unknown unit is not valid
    END_CASE
END_IF
END_FUNCTION

(* ---- FC_DL_DayOfWeekCalc.st ---- *)
(*==============================================================================
 * 组件名称 (Component)  : FC_DL_DayOfWeekCalc
 * 所属子库 (Sublibrary) : DL_Base
 * 当前版本 (Version)    : 1.0.0
 * 兼容性   (Platform)   : CODESYS 3.5 / TwinCAT 3 / 汇川 InoProShop / Machine Expert
 *                         纯 IEC 61131-3 整数运算，零库依赖，零厂商方言
 * 分类     (Category)   : 函数（FUNCTION）· 日历/星期换算 · Level 0 DL_Base 补强件
 * 功能描述 (Function)   : 年月日 → 星期几换算原子函数（ISO-8601 序：周一=1 …
 *                         周日=7）。参数域校验（年 1980..2099、月 1..12、日按
 *                         当月天数含闰年 4/100/400 判定），越界一律返回
 *                         eInvalid(0) 并置参数非法码 16#0001_0201。算法为
 *                         Sakamoto 公开算法 clean-room 实现：纯整数分段计算，
 *                         无浮点、无除零风险（除数均为非零常量 4/100/400/7）、
 *                         无循环语句（无 WHILE/REPEAT，无死锁义务，机检口径
 *                         本组件按纯分段计算豁免循环计数器审查）。
 * 开源溯源 (Origin)     : 来源标签 lgf-datetime（Siemens LGF V5.2.1 · 3.1 Date
 *                         and timer operations 章）。仅取 LGF「星期计算可拆为
 *                         独立原子 FC」的粒度结论与时间量引脚注入约定；LGF 定时
 *                         开关依赖读 CPU 本地钟，本库零全局耦合红线禁止此耦合，
 *                         日期一律由引脚注入。星期编号取 ISO-8601 周一=1，与
 *                         LGF 周日=1 惯例的差异已在规格书 §4.1 与手册显式声明
 *                         （与 GB/T 7408、MES 排产惯例一致）。核心算法为
 *                         Sakamoto 公开算法 clean-room 重写，未复制任何源码行。
 * 本文件内含       : TYPE E_DL_Weekday（星期枚举，归属 DL_Base，随本函数同文件）
 *                    FUNCTION FC_DL_DayOfWeekCalc
 * 依赖     (Depends)    : 无（纯整数运算，零 DL_ 内部依赖，可单独编译）
 * 故障码表 (Error codes) : 16#0001_0201【信息级】日期参数越界（年/月/日），
 *                          返回 eInvalid(0)；0 = 无故障。沿用 DL_Base 既有
 *                          16#0001_xxxx 段，与 VERSION.md 故障码表无冲突。
 * 红线自检 (Redline)    : R1 ✓ 零全局变量表与外部变量引用 ｜ R2 ✓ 零物理 IO 地址直写
 *                         R3 ✓ 纯 IEC 61131-3 ｜ R4 ✓ 越界防御+常量除数防除零+闰年处理
 *                         R5 ✓ 全变量中英双语同行注释 ｜ R6 不适用（无状态机，纯函数）
 *                         R7 不适用（无定时器/边沿实例）
 * 修订历史 (Revision)   :
 *   2026-11-15  v1.0.0  首版入库 · Round 05 · 泳道 B · 契约出处 ROUND_PLAN_R5 §4.1
 * 验收向量 (Acceptance) :
 *   V1 合法基准：2026-11-15 → eSunday(7)，uErrorId=0（Sakamoto 手算复核）
 *   V2 合法基准：2026-01-01 → eThursday(4)；2000-01-01 → eSaturday(6)
 *   V3 闰年边界：2024-02-29 → 合法返回（2024 为闰年，4 整除且非 100 整除）；
 *      2100-02-29 → 0001_0201（2100 为世纪非闰年，100 整除非 400 整除）；
 *      2000-02-29 → 合法返回（400 整除）
 *   V4 年越界：1979 / 2100 → eInvalid(0) + 0001_0201
 *   V5 月/日越界：uMonth=0 / 13、uDay=0 / 32、4-30、2-30 → 0001_0201
 *   V6 端年端日：1980-01-01（周三）与 2099-12-31（周四）合法返回
 *============================================================================*)

(*-----------------------------------------------------------------------------
 * 枚举: E_DL_Weekday（归属 DL_Base，与 FC_DL_DayOfWeekCalc 同文件）
 * 含义: ISO-8601 星期序，周一=1 … 周日=7；0 保留为非法/未计算值。
 *----------------------------------------------------------------------------*)
{attribute 'qualified_only'}
{attribute 'strict'}
TYPE E_DL_Weekday :
(
    eInvalid   := 0,   // 非法/未计算（Invalid），参数越界时的返回值
    eMonday    := 1,   // 周一（Monday，ISO-8601 = 1），MES 排产周首日
    eTuesday   := 2,   // 周二（Tuesday，ISO-8601 = 2）
    eWednesday := 3,   // 周三（Wednesday，ISO-8601 = 3）
    eThursday  := 4,   // 周四（Thursday，ISO-8601 = 4）
    eFriday    := 5,   // 周五（Friday，ISO-8601 = 5）
    eSaturday  := 6,   // 周六（Saturday，ISO-8601 = 6）
    eSunday    := 7    // 周日（Sunday，ISO-8601 = 7），GB/T 7408 周末日
) UINT;
END_TYPE

(*==============================================================================
 * 函数: FC_DL_DayOfWeekCalc
 * 返回值即规格引脚 eWeekday（星期几，ISO-8601 序）；非法参数返回 eInvalid(0)。
 *============================================================================*)
FUNCTION FC_DL_DayOfWeekCalc : E_DL_Weekday
VAR_INPUT
    uYear  : UINT;    // 年份（Year）[年]，有效域 1980..2099，越界返回 eInvalid
    uMonth : USINT;   // 月（Month）[月]，有效域 1..12，越界返回 eInvalid
    uDay   : USINT;   // 日（Day）[日]，有效域 1..当月天数（含闰年 2 月 29 日），越界返回 eInvalid
END_VAR
VAR_OUTPUT
    uErrorId : UDINT; // 参数非法码（Error code）：16#0001_0201 = 日期越界；0 = 合法
END_VAR
VAR
    _nY    : DINT;    // 算法内部年（1~2 月按 Sakamoto 惯例回退一年）[年]
    _nT    : DINT;    // Sakamoto 月修正表值（Month offset of Sakamoto table）
    _nWd   : DINT;    // 星期原始值（Raw weekday）0=周日..6=周六
    _nIso  : DINT;    // ISO-8601 星期（ISO weekday）1=周一..7=周日
    _nDim  : DINT;    // 当月天数（Days in month）28..31
    _bLeap : BOOL;    // 闰年标志（Leap year flag），判定规则 4/100/400
END_VAR

// 段 0｜出口默认值先赋（公约 0.8 精神：防御路径之前），越界路径直接沿用此默认
FC_DL_DayOfWeekCalc := E_DL_Weekday.eInvalid;  // 默认返回非法枚举
uErrorId := 16#0001_0201;                      // 默认携带参数越界码（信息级）

// 段 1｜参数域校验：年（规格 §4.1 固定域 1980..2099）
IF (uYear < 1980) OR (uYear > 2099) THEN
    RETURN;                                    // 年越界：保持默认 eInvalid + 0001_0201
END_IF

// 段 2｜参数域校验：月
IF (uMonth < 1) OR (uMonth > 12) THEN
    RETURN;                                    // 月越界：保持默认
END_IF

// 段 3｜闰年判定（4/100/400 三段规则：世纪年须 400 整除）
_nY    := uYear;                               // UINT → DINT 隐式扩宽，无精度损失
_bLeap := (( (_nY MOD 4) = 0) AND ( (_nY MOD 100) <> 0))
       OR ( (_nY MOD 400) = 0);                // 整除判定用 MOD，除数为非零常量，无除零风险

// 段 4｜当月天数与日校验（CASE 兜底分支为不可达防御位，R6 精神）
CASE uMonth OF
    1, 3, 5, 7, 8, 10, 12:  _nDim := 31;       // 大月 31 天
    4, 6, 9, 11:            _nDim := 30;       // 小月 30 天
    2:                                          // 二月按闰年分档
        IF _bLeap THEN
            _nDim := 29;                       // 闰年二月 29 天
        ELSE
            _nDim := 28;                       // 平年二月 28 天
        END_IF
    ELSE
        _nDim := 0;                            // 不可达防御位（月已校验 1..12）
END_CASE
IF (uDay < 1) OR (uDay > _nDim) THEN
    RETURN;                                    // 日越界（含平年 2-29、小月 31 日）：保持默认
END_IF

// 段 5｜Sakamoto 分段计算：1~2 月按惯例回退一年再取月修正表
IF uMonth < 3 THEN
    _nY := _nY - 1;                            // 1~2 月回退一年（Sakamoto 惯例）
END_IF
CASE uMonth OF
    1:  _nT := 0;                              // 月修正表（Sakamoto table，一月）
    2:  _nT := 3;                              // 二月
    3:  _nT := 2;                              // 三月
    4:  _nT := 5;                              // 四月
    5:  _nT := 0;                              // 五月
    6:  _nT := 3;                              // 六月
    7:  _nT := 5;                              // 七月
    8:  _nT := 1;                              // 八月
    9:  _nT := 4;                              // 九月
    10: _nT := 6;                              // 十月
    11: _nT := 2;                              // 十一月
    12: _nT := 4;                              // 十二月
    ELSE
        _nT := 0;                              // 不可达防御位（月已校验 1..12）
END_CASE

// 段 6｜星期合成：纯整数四则 + 常量模 7，结果域 0=周日..6=周六
_nWd := (_nY + (_nY / 4) - (_nY / 100) + (_nY / 400) + _nT + uDay) MOD 7;
//  说明：除数 4/100/400/7 均为非零常量，DINT 正数域整除，无除零风险（R4）

// 段 7｜ISO-8601 换算：0(周日)→7，1..6(周一..周六)→1..6
_nIso := ((_nWd + 6) MOD 7) + 1;

// 段 8｜映射到枚举（strict 枚举不允许整型直赋，显式 CASE 映射）
CASE _nIso OF
    1: FC_DL_DayOfWeekCalc := E_DL_Weekday.eMonday;     // 周一
    2: FC_DL_DayOfWeekCalc := E_DL_Weekday.eTuesday;    // 周二
    3: FC_DL_DayOfWeekCalc := E_DL_Weekday.eWednesday;  // 周三
    4: FC_DL_DayOfWeekCalc := E_DL_Weekday.eThursday;   // 周四
    5: FC_DL_DayOfWeekCalc := E_DL_Weekday.eFriday;     // 周五
    6: FC_DL_DayOfWeekCalc := E_DL_Weekday.eSaturday;   // 周六
    7: FC_DL_DayOfWeekCalc := E_DL_Weekday.eSunday;     // 周日
    ELSE
        FC_DL_DayOfWeekCalc := E_DL_Weekday.eInvalid;   // 不可达防御位（_nIso 恒 1..7）
END_CASE

uErrorId := 16#0000_0000;                      // 合法路径清码

END_FUNCTION
